Universal Robots URScript: jerry_new_robot_1.script

def Machining2():
  # Default parameters:
  global speed_ms = 0.3
  global speed_rads = 0.75
  global accel_mss = 3
  global accel_radss = 1.2
  global blend_radius_m = 0.001

  # Add subprograms here
  # Start of main program
  # Program generated by RoboDK v5.6.8 for UR10e on 15/12/2023 14:31:05
  # Using nominal kinematics.
  blend_radius_m = 0.001
  speed_ms = 0.01
  # set_reference(p[0.405000, -0.105000, 0.010000, 0.000000, 0.000000, 0.000000])
  set_tcp(p[0.000000, 0.000000, 0.252000, 0.000000, 0.000000, 0.000000])
  # Show Tool
  movej([0.286818, -1.328197, -2.476759, -0.907433, 1.570796, 1.857614],accel_radss,speed_rads,0,blend_radius_m)
  movel([0.286818, -1.380785, -2.509088, -0.822516, 1.570796, 1.857614],accel_mss,speed_ms,0,blend_radius_m)
  speed_ms = 0.01
  movel([0.286818, -1.403946, -2.521184, -0.787258, 1.570796, 1.857614],accel_mss,speed_ms,0,blend_radius_m)
  speed_ms = 0.003
  movel([0.286818, -1.412952, -2.525590, -0.773847, 1.570796, 1.857614],accel_mss,speed_ms,0,blend_radius_m)
  speed_ms = 0.007
  movel([0.278957, -1.415271, -2.523827, -0.773292, 1.570796, 1.849754],accel_mss,speed_ms,0,blend_radius_m)
  movel([0.277121, -1.413155, -2.525436, -0.773798, 1.570796, 1.847918],accel_mss,speed_ms,0,blend_radius_m)
  movel([0.275274, -1.411040, -2.527038, -0.774311, 1.570796, 1.846071],accel_mss,speed_ms,0,blend_radius_m)
  movel([0.275922, -1.409907, -2.527894, -0.774588, 1.570796, 1.846719],accel_mss,speed_ms,0,blend_radius_m)
  movel([0.276572, -1.408773, -2.528749, -0.774868, 1.570796, 1.847368],accel_mss,speed_ms,0,blend_radius_m)
  movel([0.275763, -1.408648, -2.528842, -0.774898, 1.570796, 1.846559],accel_mss,speed_ms,0,blend_radius_m)
  movel([0.268969, -1.407825, -2.529461, -0.775102, 1.570796, 1.839766],accel_mss,speed_ms,0,blend_radius_m)
  movel([0.266583, -1.407546, -2.529671, -0.775172, 1.570796, 1.837380],accel_mss,speed_ms,0,blend_radius_m)
  movel([0.265501, -1.407413, -2.529771, -0.775205, 1.570796, 1.836297],accel_mss,speed_ms,0,blend_radius_m)
  movel([0.264422, -1.407272, -2.529877, -0.775240, 1.570796, 1.835218],accel_mss,speed_ms,0,blend_radius_m)
  movel([0.263348, -1.407121, -2.529990, -0.775278, 1.570796, 1.834144],accel_mss,speed_ms,0,blend_radius_m)
  movel([0.262516, -1.406998, -2.530083, -0.775309, 1.570796, 1.833312],accel_mss,speed_ms,0,blend_radius_m)
  movel([0.261691, -1.406866, -2.530182, -0.775342, 1.570796, 1.832487],accel_mss,speed_ms,0,blend_radius_m)
  movel([0.260873, -1.406721, -2.530290, -0.775378, 1.570796, 1.831670],accel_mss,speed_ms,0,blend_radius_m)
  movel([0.260123, -1.406582, -2.530395, -0.775413, 1.570796, 1.830919],accel_mss,speed_ms,0,blend_radius_m)
  movel([0.259383, -1.406429, -2.530509, -0.775451, 1.570796, 1.830179],accel_mss,speed_ms,0,blend_radius_m)
  movel([0.258650, -1.406263, -2.530633, -0.775493, 1.570796, 1.829447],accel_mss,speed_ms,0,blend_radius_m)
  movel([0.257946, -1.406092, -2.530761, -0.775535, 1.570796, 1.828742],accel_mss,speed_ms,0,blend_radius_m)
  movel([0.257255, -1.405904, -2.530902, -0.775583, 1.570796, 1.828051],accel_mss,speed_ms,0,blend_radius_m)
  movel([0.256572, -1.405700, -2.531055, -0.775634, 1.570796, 1.827368],accel_mss,speed_ms,0,blend_radius_m)
  movel([0.255900, -1.405481, -2.531218, -0.775689, 1.570796, 1.826696],accel_mss,speed_ms,0,blend_radius_m)
  movel([0.255241, -1.405247, -2.531394, -0.775748, 1.570796, 1.826037],accel_mss,speed_ms,0,blend_radius_m)
  movel([0.254785, -1.405071, -2.531525, -0.775793, 1.570796, 1.825581],accel_mss,speed_ms,0,blend_radius_m)
  movel([0.254341, -1.404877, -2.531670, -0.775842, 1.570796, 1.825137],accel_mss,speed_ms,0,blend_radius_m)
  movel([0.253906, -1.404672, -2.531824, -0.775894, 1.570796, 1.824702],accel_mss,speed_ms,0,blend_radius_m)
  movel([0.253487, -1.404450, -2.531989, -0.775950, 1.570796, 1.824283],accel_mss,speed_ms,0,blend_radius_m)
  movel([0.253079, -1.404213, -2.532166, -0.776010, 1.570796, 1.823875],accel_mss,speed_ms,0,blend_radius_m)
  movel([0.252685, -1.403964, -2.532352, -0.776073, 1.570796, 1.823481],accel_mss,speed_ms,0,blend_radius_m)
  movel([0.252356, -1.403735, -2.532523, -0.776131, 1.570796, 1.823152],accel_mss,speed_ms,0,blend_radius_m)
  movel([0.252040, -1.403492, -2.532704, -0.776193, 1.570796, 1.822837],accel_mss,speed_ms,0,blend_radius_m)
  movel([0.251741, -1.403234, -2.532896, -0.776259, 1.570796, 1.822538],accel_mss,speed_ms,0,blend_radius_m)
  movel([0.251455, -1.402963, -2.533098, -0.776328, 1.570796, 1.822252],accel_mss,speed_ms,0,blend_radius_m)
  movel([0.251184, -1.402679, -2.533309, -0.776401, 1.570796, 1.821980],accel_mss,speed_ms,0,blend_radius_m)
  movel([0.250929, -1.402382, -2.533530, -0.776477, 1.570796, 1.821725],accel_mss,speed_ms,0,blend_radius_m)
  movel([0.250744, -1.402139, -2.533711, -0.776540, 1.570796, 1.821540],accel_mss,speed_ms,0,blend_radius_m)
  movel([0.250570, -1.401887, -2.533898, -0.776604, 1.570796, 1.821366],accel_mss,speed_ms,0,blend_radius_m)
  movel([0.250413, -1.401623, -2.534094, -0.776672, 1.570796, 1.821209],accel_mss,speed_ms,0,blend_radius_m)
  movel([0.250269, -1.401348, -2.534298, -0.776743, 1.570796, 1.821066],accel_mss,speed_ms,0,blend_radius_m)
  movel([0.250142, -1.401063, -2.534509, -0.776817, 1.570796, 1.820938],accel_mss,speed_ms,0,blend_radius_m)
  movel([0.250030, -1.400772, -2.534725, -0.776892, 1.570796, 1.820826],accel_mss,speed_ms,0,blend_radius_m)
  movel([0.249933, -1.400468, -2.534950, -0.776970, 1.570796, 1.820729],accel_mss,speed_ms,0,blend_radius_m)
  movel([0.249858, -1.400178, -2.535165, -0.777046, 1.570796, 1.820655],accel_mss,speed_ms,0,blend_radius_m)
  movel([0.249800, -1.399877, -2.535388, -0.777124, 1.570796, 1.820596],accel_mss,speed_ms,0,blend_radius_m)
  movel([0.249762, -1.399567, -2.535617, -0.777205, 1.570796, 1.820559],accel_mss,speed_ms,0,blend_radius_m)
  movel([0.249742, -1.399250, -2.535851, -0.777287, 1.570796, 1.820538],accel_mss,speed_ms,0,blend_radius_m)
  movel([0.249739, -1.398896, -2.536113, -0.777380, 1.570796, 1.820535],accel_mss,speed_ms,0,blend_radius_m)
  movel([0.249750, -1.398537, -2.536378, -0.777474, 1.570796, 1.820546],accel_mss,speed_ms,0,blend_radius_m)
  movel([0.249777, -1.398172, -2.536647, -0.777570, 1.570796, 1.820573],accel_mss,speed_ms,0,blend_radius_m)
  movel([0.249818, -1.397802, -2.536920, -0.777667, 1.570796, 1.820614],accel_mss,speed_ms,0,blend_radius_m)
  movel([0.249880, -1.397415, -2.537205, -0.777769, 1.570796, 1.820676],accel_mss,speed_ms,0,blend_radius_m)
  movel([0.249952, -1.397029, -2.537490, -0.777871, 1.570796, 1.820749],accel_mss,speed_ms,0,blend_radius_m)
  movel([0.250043, -1.396635, -2.537779, -0.777975, 1.570796, 1.820839],accel_mss,speed_ms,0,blend_radius_m)
  movel([0.250147, -1.396242, -2.538068, -0.778079, 1.570796, 1.820943],accel_mss,speed_ms,0,blend_radius_m)
  movel([0.250264, -1.395857, -2.538351, -0.778181, 1.570796, 1.821061],accel_mss,speed_ms,0,blend_radius_m)
  movel([0.250398, -1.395471, -2.538634, -0.778284, 1.570796, 1.821194],accel_mss,speed_ms,0,blend_radius_m)
  movel([0.250547, -1.395084, -2.538918, -0.778387, 1.570796, 1.821344],accel_mss,speed_ms,0,blend_radius_m)
  movel([0.250711, -1.394696, -2.539203, -0.778491, 1.570796, 1.821507],accel_mss,speed_ms,0,blend_radius_m)
  movel([0.250904, -1.394272, -2.539513, -0.778604, 1.570796, 1.821701],accel_mss,speed_ms,0,blend_radius_m)
  movel([0.251110, -1.393847, -2.539824, -0.778719, 1.570796, 1.821906],accel_mss,speed_ms,0,blend_radius_m)
  movel([0.251326, -1.393423, -2.540133, -0.778832, 1.570796, 1.822123],accel_mss,speed_ms,0,blend_radius_m)
  movel([0.251379, -1.393339, -2.540195, -0.778855, 1.570796, 1.822175],accel_mss,speed_ms,0,blend_radius_m)
  movel([0.251441, -1.393255, -2.540256, -0.778878, 1.570796, 1.822237],accel_mss,speed_ms,0,blend_radius_m)
  movel([0.251514, -1.393178, -2.540313, -0.778899, 1.570796, 1.822310],accel_mss,speed_ms,0,blend_radius_m)
  movel([0.251592, -1.393106, -2.540365, -0.778918, 1.570796, 1.822389],accel_mss,speed_ms,0,blend_radius_m)
  movel([0.251680, -1.393042, -2.540412, -0.778935, 1.570796, 1.822476],accel_mss,speed_ms,0,blend_radius_m)
  movel([0.251772, -1.392987, -2.540452, -0.778950, 1.570796, 1.822568],accel_mss,speed_ms,0,blend_radius_m)
  movel([0.251894, -1.392931, -2.540493, -0.778965, 1.570796, 1.822690],accel_mss,speed_ms,0,blend_radius_m)
  movel([0.252016, -1.392887, -2.540525, -0.778977, 1.570796, 1.822813],accel_mss,speed_ms,0,blend_radius_m)
  movel([0.252140, -1.392857, -2.540547, -0.778985, 1.570796, 1.822936],accel_mss,speed_ms,0,blend_radius_m)
  movel([0.252259, -1.392843, -2.540557, -0.778989, 1.570796, 1.823055],accel_mss,speed_ms,0,blend_radius_m)
  movel([0.252371, -1.392844, -2.540556, -0.778989, 1.570796, 1.823167],accel_mss,speed_ms,0,blend_radius_m)
  movel([0.252874, -1.392895, -2.540519, -0.778975, 1.570796, 1.823670],accel_mss,speed_ms,0,blend_radius_m)
  movel([0.253372, -1.392952, -2.540477, -0.778959, 1.570796, 1.824168],accel_mss,speed_ms,0,blend_radius_m)
  movel([0.253866, -1.393017, -2.540430, -0.778942, 1.570796, 1.824662],accel_mss,speed_ms,0,blend_radius_m)
  movel([0.254596, -1.393123, -2.540352, -0.778913, 1.570796, 1.825392],accel_mss,speed_ms,0,blend_radius_m)
  movel([0.254793, -1.392422, -2.540864, -0.779103, 1.570796, 1.825589],accel_mss,speed_ms,0,blend_radius_m)
  movel([0.254989, -1.391722, -2.541374, -0.779293, 1.570796, 1.825785],accel_mss,speed_ms,0,blend_radius_m)
  movel([0.238692, -1.394040, -2.539683, -0.778667, 1.570796, 1.809488],accel_mss,speed_ms,0,blend_radius_m)
  movel([0.229160, -1.395492, -2.538618, -0.778278, 1.570796, 1.799956],accel_mss,speed_ms,0,blend_radius_m)
  movel([0.227094, -1.395812, -2.538384, -0.778193, 1.570796, 1.797890],accel_mss,speed_ms,0,blend_radius_m)
  movel([0.225031, -1.396124, -2.538155, -0.778110, 1.570796, 1.795827],accel_mss,speed_ms,0,blend_radius_m)
  movel([0.222484, -1.396503, -2.537876, -0.778010, 1.570796, 1.793281],accel_mss,speed_ms,0,blend_radius_m)
  movel([0.222392, -1.396509, -2.537872, -0.778008, 1.570796, 1.793189],accel_mss,speed_ms,0,blend_radius_m)
  movel([0.222306, -1.396503, -2.537876, -0.778010, 1.570796, 1.793102],accel_mss,speed_ms,0,blend_radius_m)
  movel([0.222225, -1.396485, -2.537890, -0.778014, 1.570796, 1.793021],accel_mss,speed_ms,0,blend_radius_m)
  movel([0.222156, -1.396453, -2.537913, -0.778023, 1.570796, 1.792952],accel_mss,speed_ms,0,blend_radius_m)
  movel([0.222108, -1.396419, -2.537938, -0.778032, 1.570796, 1.792904],accel_mss,speed_ms,0,blend_radius_m)
  movel([0.222070, -1.396378, -2.537968, -0.778043, 1.570796, 1.792867],accel_mss,speed_ms,0,blend_radius_m)
  movel([0.222044, -1.396328, -2.538005, -0.778056, 1.570796, 1.792841],accel_mss,speed_ms,0,blend_radius_m)
  movel([0.222025, -1.396269, -2.538048, -0.778072, 1.570796, 1.792821],accel_mss,speed_ms,0,blend_radius_m)
  movel([0.222016, -1.396204, -2.538096, -0.778089, 1.570796, 1.792812],accel_mss,speed_ms,0,blend_radius_m)
  movel([0.222016, -1.396138, -2.538144, -0.778106, 1.570796, 1.792813],accel_mss,speed_ms,0,blend_radius_m)
  movel([0.222040, -1.395960, -2.538275, -0.778154, 1.570796, 1.792836],accel_mss,speed_ms,0,blend_radius_m)
  movel([0.222075, -1.395781, -2.538407, -0.778201, 1.570796, 1.792872],accel_mss,speed_ms,0,blend_radius_m)
  movel([0.222291, -1.394877, -2.539069, -0.778442, 1.570796, 1.793087],accel_mss,speed_ms,0,blend_radius_m)
  movel([0.222650, -1.393424, -2.540133, -0.778832, 1.570796, 1.793446],accel_mss,speed_ms,0,blend_radius_m)
  movel([0.212968, -1.395043, -2.538948, -0.778398, 1.570796, 1.783765],accel_mss,speed_ms,0,blend_radius_m)
  movel([0.203286, -1.396738, -2.537704, -0.777948, 1.570796, 1.774082],accel_mss,speed_ms,0,blend_radius_m)
  movel([0.203152, -1.397328, -2.537269, -0.777792, 1.570796, 1.773949],accel_mss,speed_ms,0,blend_radius_m)
  movel([0.203019, -1.397918, -2.536835, -0.777636, 1.570796, 1.773815],accel_mss,speed_ms,0,blend_radius_m)
  movel([0.186235, -1.401026, -2.534537, -0.776826, 1.570796, 1.757031],accel_mss,speed_ms,0,blend_radius_m)
  movel([0.169460, -1.404353, -2.532062, -0.775974, 1.570796, 1.740256],accel_mss,speed_ms,0,blend_radius_m)
  movel([0.168502, -1.404999, -2.531579, -0.775811, 1.570796, 1.739298],accel_mss,speed_ms,0,blend_radius_m)
  movel([0.168210, -1.405190, -2.531436, -0.775763, 1.570796, 1.739006],accel_mss,speed_ms,0,blend_radius_m)
  movel([0.167917, -1.405378, -2.531296, -0.775715, 1.570796, 1.738713],accel_mss,speed_ms,0,blend_radius_m)
  movel([0.167618, -1.405559, -2.531161, -0.775670, 1.570796, 1.738414],accel_mss,speed_ms,0,blend_radius_m)
  movel([0.167135, -1.405842, -2.530948, -0.775598, 1.570796, 1.737931],accel_mss,speed_ms,0,blend_radius_m)
  movel([0.166648, -1.406110, -2.530748, -0.775531, 1.570796, 1.737444],accel_mss,speed_ms,0,blend_radius_m)
  movel([0.166146, -1.406376, -2.530549, -0.775464, 1.570796, 1.736942],accel_mss,speed_ms,0,blend_radius_m)
  movel([0.165641, -1.406626, -2.530362, -0.775402, 1.570796, 1.736437],accel_mss,speed_ms,0,blend_radius_m)
  movel([0.165143, -1.406860, -2.530186, -0.775343, 1.570796, 1.735939],accel_mss,speed_ms,0,blend_radius_m)
  movel([0.164644, -1.407079, -2.530022, -0.775288, 1.570796, 1.735440],accel_mss,speed_ms,0,blend_radius_m)
  movel([0.164316, -1.407211, -2.529922, -0.775255, 1.570796, 1.735113],accel_mss,speed_ms,0,blend_radius_m)
  movel([0.163987, -1.407330, -2.529833, -0.775226, 1.570796, 1.734783],accel_mss,speed_ms,0,blend_radius_m)
  movel([0.163661, -1.407432, -2.529756, -0.775200, 1.570796, 1.734457],accel_mss,speed_ms,0,blend_radius_m)
  movel([0.162882, -1.407653, -2.529590, -0.775145, 1.570796, 1.733678],accel_mss,speed_ms,0,blend_radius_m)
  movel([0.162106, -1.407860, -2.529435, -0.775094, 1.570796, 1.732902],accel_mss,speed_ms,0,blend_radius_m)
  movel([0.161310, -1.408059, -2.529285, -0.775044, 1.570796, 1.732107],accel_mss,speed_ms,0,blend_radius_m)
  movel([0.160517, -1.408252, -2.529140, -0.774996, 1.570796, 1.731313],accel_mss,speed_ms,0,blend_radius_m)
  movel([0.160414, -1.408270, -2.529127, -0.774992, 1.570796, 1.731210],accel_mss,speed_ms,0,blend_radius_m)
  movel([0.160319, -1.408272, -2.529125, -0.774992, 1.570796, 1.731115],accel_mss,speed_ms,0,blend_radius_m)
  movel([0.160228, -1.408261, -2.529134, -0.774994, 1.570796, 1.731025],accel_mss,speed_ms,0,blend_radius_m)
  movel([0.160150, -1.408233, -2.529155, -0.775001, 1.570796, 1.730946],accel_mss,speed_ms,0,blend_radius_m)
  movel([0.160120, -1.408213, -2.529170, -0.775006, 1.570796, 1.730916],accel_mss,speed_ms,0,blend_radius_m)
  movel([0.160100, -1.408185, -2.529191, -0.775013, 1.570796, 1.730896],accel_mss,speed_ms,0,blend_radius_m)
  movel([0.160090, -1.408151, -2.529216, -0.775021, 1.570796, 1.730887],accel_mss,speed_ms,0,blend_radius_m)
  movel([0.160090, -1.408113, -2.529245, -0.775031, 1.570796, 1.730887],accel_mss,speed_ms,0,blend_radius_m)
  movel([0.160497, -1.405621, -2.531114, -0.775654, 1.570796, 1.731293],accel_mss,speed_ms,0,blend_radius_m)
  movel([0.160790, -1.403859, -2.532430, -0.776100, 1.570796, 1.731586],accel_mss,speed_ms,0,blend_radius_m)
  movel([0.161094, -1.402089, -2.533748, -0.776552, 1.570796, 1.731890],accel_mss,speed_ms,0,blend_radius_m)
  movel([0.162202, -1.395764, -2.538419, -0.778206, 1.570796, 1.732999],accel_mss,speed_ms,0,blend_radius_m)
  movel([0.164448, -1.383126, -2.547582, -0.781681, 1.570796, 1.735244],accel_mss,speed_ms,0,blend_radius_m)
  movel([0.164830, -1.383043, -2.547641, -0.781705, 1.570796, 1.735626],accel_mss,speed_ms,0,blend_radius_m)
  movel([0.165050, -1.382984, -2.547683, -0.781721, 1.570796, 1.735846],accel_mss,speed_ms,0,blend_radius_m)
  movel([0.165159, -1.382921, -2.547729, -0.781739, 1.570796, 1.735955],accel_mss,speed_ms,0,blend_radius_m)
  movel([0.165225, -1.382825, -2.547797, -0.781767, 1.570796, 1.736022],accel_mss,speed_ms,0,blend_radius_m)
  movel([0.165270, -1.382649, -2.547923, -0.781817, 1.570796, 1.736066],accel_mss,speed_ms,0,blend_radius_m)
  movel([0.165294, -1.382556, -2.547990, -0.781843, 1.570796, 1.736090],accel_mss,speed_ms,0,blend_radius_m)
  movel([0.165328, -1.382461, -2.548058, -0.781870, 1.570796, 1.736124],accel_mss,speed_ms,0,blend_radius_m)
  movel([0.165349, -1.382421, -2.548086, -0.781882, 1.570796, 1.736145],accel_mss,speed_ms,0,blend_radius_m)
  movel([0.165379, -1.382383, -2.548113, -0.781893, 1.570796, 1.736176],accel_mss,speed_ms,0,blend_radius_m)
  movel([0.165418, -1.382352, -2.548136, -0.781902, 1.570796, 1.736214],accel_mss,speed_ms,0,blend_radius_m)
  movel([0.165499, -1.382303, -2.548171, -0.781915, 1.570796, 1.736295],accel_mss,speed_ms,0,blend_radius_m)
  movel([0.165585, -1.382265, -2.548198, -0.781926, 1.570796, 1.736381],accel_mss,speed_ms,0,blend_radius_m)
  movel([0.166012, -1.382128, -2.548296, -0.781965, 1.570796, 1.736808],accel_mss,speed_ms,0,blend_radius_m)
  movel([0.166274, -1.382054, -2.548348, -0.781986, 1.570796, 1.737070],accel_mss,speed_ms,0,blend_radius_m)
  movel([0.166534, -1.381992, -2.548393, -0.782004, 1.570796, 1.737330],accel_mss,speed_ms,0,blend_radius_m)
  movel([0.166792, -1.381940, -2.548430, -0.782019, 1.570796, 1.737589],accel_mss,speed_ms,0,blend_radius_m)
  movel([0.167305, -1.381853, -2.548492, -0.782044, 1.570796, 1.738102],accel_mss,speed_ms,0,blend_radius_m)
  movel([0.167813, -1.381783, -2.548542, -0.782064, 1.570796, 1.738609],accel_mss,speed_ms,0,blend_radius_m)
  movel([0.168346, -1.381724, -2.548584, -0.782081, 1.570796, 1.739143],accel_mss,speed_ms,0,blend_radius_m)
  movel([0.168877, -1.381683, -2.548614, -0.782092, 1.570796, 1.739673],accel_mss,speed_ms,0,blend_radius_m)
  movel([0.169191, -1.381665, -2.548626, -0.782098, 1.570796, 1.739987],accel_mss,speed_ms,0,blend_radius_m)
  movel([0.169501, -1.381659, -2.548631, -0.782099, 1.570796, 1.740297],accel_mss,speed_ms,0,blend_radius_m)
  movel([0.169807, -1.381660, -2.548630, -0.782099, 1.570796, 1.740603],accel_mss,speed_ms,0,blend_radius_m)
  movel([0.170079, -1.381669, -2.548624, -0.782097, 1.570796, 1.740875],accel_mss,speed_ms,0,blend_radius_m)
  movel([0.170344, -1.381689, -2.548609, -0.782091, 1.570796, 1.741141],accel_mss,speed_ms,0,blend_radius_m)
  movel([0.170606, -1.381717, -2.548590, -0.782083, 1.570796, 1.741402],accel_mss,speed_ms,0,blend_radius_m)
  movel([0.171068, -1.381785, -2.548541, -0.782063, 1.570796, 1.741865],accel_mss,speed_ms,0,blend_radius_m)
  movel([0.171524, -1.381865, -2.548483, -0.782040, 1.570796, 1.742320],accel_mss,speed_ms,0,blend_radius_m)
  movel([0.171974, -1.381962, -2.548415, -0.782013, 1.570796, 1.742770],accel_mss,speed_ms,0,blend_radius_m)
  movel([0.172412, -1.382071, -2.548336, -0.781982, 1.570796, 1.743208],accel_mss,speed_ms,0,blend_radius_m)
  movel([0.172651, -1.382141, -2.548286, -0.781961, 1.570796, 1.743447],accel_mss,speed_ms,0,blend_radius_m)
  movel([0.172886, -1.382221, -2.548229, -0.781939, 1.570796, 1.743682],accel_mss,speed_ms,0,blend_radius_m)
  movel([0.173112, -1.382309, -2.548166, -0.781914, 1.570796, 1.743908],accel_mss,speed_ms,0,blend_radius_m)
  movel([0.173605, -1.382514, -2.548020, -0.781855, 1.570796, 1.744401],accel_mss,speed_ms,0,blend_radius_m)
  movel([0.190906, -1.378978, -2.550540, -0.782871, 1.570796, 1.761702],accel_mss,speed_ms,0,blend_radius_m)
  movel([0.208219, -1.375672, -2.552880, -0.783837, 1.570796, 1.779015],accel_mss,speed_ms,0,blend_radius_m)
  movel([0.208066, -1.376337, -2.552411, -0.783642, 1.570796, 1.778862],accel_mss,speed_ms,0,blend_radius_m)
  movel([0.207913, -1.377000, -2.551942, -0.783447, 1.570796, 1.778709],accel_mss,speed_ms,0,blend_radius_m)
  movel([0.212684, -1.376133, -2.552555, -0.783702, 1.570796, 1.783480],accel_mss,speed_ms,0,blend_radius_m)
  movel([0.217469, -1.375223, -2.553196, -0.783969, 1.570796, 1.788265],accel_mss,speed_ms,0,blend_radius_m)
  movel([0.217297, -1.374328, -2.553827, -0.784234, 1.570796, 1.788093],accel_mss,speed_ms,0,blend_radius_m)
  movel([0.217253, -1.374069, -2.554009, -0.784311, 1.570796, 1.788049],accel_mss,speed_ms,0,blend_radius_m)
  movel([0.217221, -1.373807, -2.554194, -0.784389, 1.570796, 1.788017],accel_mss,speed_ms,0,blend_radius_m)
  movel([0.217200, -1.373555, -2.554371, -0.784464, 1.570796, 1.787996],accel_mss,speed_ms,0,blend_radius_m)
  movel([0.217190, -1.373298, -2.554551, -0.784540, 1.570796, 1.787986],accel_mss,speed_ms,0,blend_radius_m)
  movel([0.217192, -1.373038, -2.554734, -0.784618, 1.570796, 1.787988],accel_mss,speed_ms,0,blend_radius_m)
  movel([0.217206, -1.372767, -2.554924, -0.784699, 1.570796, 1.788002],accel_mss,speed_ms,0,blend_radius_m)
  movel([0.217230, -1.372493, -2.555115, -0.784780, 1.570796, 1.788026],accel_mss,speed_ms,0,blend_radius_m)
  movel([0.217264, -1.372216, -2.555310, -0.784863, 1.570796, 1.788060],accel_mss,speed_ms,0,blend_radius_m)
  movel([0.217314, -1.371908, -2.555526, -0.784955, 1.570796, 1.788111],accel_mss,speed_ms,0,blend_radius_m)
  movel([0.217375, -1.371598, -2.555742, -0.785048, 1.570796, 1.788171],accel_mss,speed_ms,0,blend_radius_m)
  movel([0.217443, -1.371287, -2.555960, -0.785142, 1.570796, 1.788239],accel_mss,speed_ms,0,blend_radius_m)
  movel([0.217532, -1.370935, -2.556206, -0.785248, 1.570796, 1.788328],accel_mss,speed_ms,0,blend_radius_m)
  movel([0.217633, -1.370581, -2.556453, -0.785354, 1.570796, 1.788429],accel_mss,speed_ms,0,blend_radius_m)
  movel([0.217749, -1.370225, -2.556702, -0.785462, 1.570796, 1.788545],accel_mss,speed_ms,0,blend_radius_m)
  movel([0.217869, -1.369901, -2.556928, -0.785560, 1.570796, 1.788665],accel_mss,speed_ms,0,blend_radius_m)
  movel([0.218003, -1.369575, -2.557155, -0.785658, 1.570796, 1.788799],accel_mss,speed_ms,0,blend_radius_m)
  movel([0.218156, -1.369250, -2.557382, -0.785757, 1.570796, 1.788952],accel_mss,speed_ms,0,blend_radius_m)
  movel([0.218328, -1.368913, -2.557617, -0.785859, 1.570796, 1.789124],accel_mss,speed_ms,0,blend_radius_m)
  movel([0.218513, -1.368579, -2.557849, -0.785961, 1.570796, 1.789309],accel_mss,speed_ms,0,blend_radius_m)
  movel([0.218715, -1.368245, -2.558082, -0.786063, 1.570796, 1.789511],accel_mss,speed_ms,0,blend_radius_m)
  movel([0.218964, -1.367856, -2.558351, -0.786181, 1.570796, 1.789761],accel_mss,speed_ms,0,blend_radius_m)
  movel([0.219223, -1.367471, -2.558619, -0.786299, 1.570796, 1.790019],accel_mss,speed_ms,0,blend_radius_m)
  movel([0.219493, -1.367087, -2.558885, -0.786417, 1.570796, 1.790290],accel_mss,speed_ms,0,blend_radius_m)
  movel([0.220268, -1.366008, -2.559633, -0.786748, 1.570796, 1.791064],accel_mss,speed_ms,0,blend_radius_m)
  movel([0.218931, -1.366247, -2.559468, -0.786674, 1.570796, 1.789727],accel_mss,speed_ms,0,blend_radius_m)
  movel([0.217591, -1.366488, -2.559301, -0.786601, 1.570796, 1.788387],accel_mss,speed_ms,0,blend_radius_m)
  movel([0.217739, -1.365869, -2.559729, -0.786791, 1.570796, 1.788535],accel_mss,speed_ms,0,blend_radius_m)
  movel([0.217888, -1.365249, -2.560158, -0.786982, 1.570796, 1.788684],accel_mss,speed_ms,0,blend_radius_m)
  movel([0.213855, -1.365983, -2.559650, -0.786756, 1.570796, 1.784651],accel_mss,speed_ms,0,blend_radius_m)
  movel([0.209822, -1.366730, -2.559133, -0.786526, 1.570796, 1.780618],accel_mss,speed_ms,0,blend_radius_m)
  movel([0.209666, -1.367404, -2.558666, -0.786320, 1.570796, 1.780462],accel_mss,speed_ms,0,blend_radius_m)
  movel([0.209510, -1.368076, -2.558199, -0.786114, 1.570796, 1.780306],accel_mss,speed_ms,0,blend_radius_m)
  movel([0.191959, -1.371470, -2.555832, -0.785087, 1.570796, 1.762755],accel_mss,speed_ms,0,blend_radius_m)
  movel([0.174421, -1.375101, -2.553282, -0.784005, 1.570796, 1.745218],accel_mss,speed_ms,0,blend_radius_m)
  movel([0.173235, -1.375825, -2.552772, -0.783792, 1.570796, 1.744031],accel_mss,speed_ms,0,blend_radius_m)
  movel([0.172826, -1.376067, -2.552601, -0.783721, 1.570796, 1.743622],accel_mss,speed_ms,0,blend_radius_m)
  movel([0.172415, -1.376300, -2.552436, -0.783652, 1.570796, 1.743211],accel_mss,speed_ms,0,blend_radius_m)
  movel([0.172001, -1.376524, -2.552278, -0.783587, 1.570796, 1.742797],accel_mss,speed_ms,0,blend_radius_m)
  movel([0.171584, -1.376736, -2.552129, -0.783525, 1.570796, 1.742381],accel_mss,speed_ms,0,blend_radius_m)
  movel([0.171160, -1.376943, -2.551982, -0.783464, 1.570796, 1.741956],accel_mss,speed_ms,0,blend_radius_m)
  movel([0.170730, -1.377139, -2.551844, -0.783407, 1.570796, 1.741527],accel_mss,speed_ms,0,blend_radius_m)
  movel([0.170303, -1.377326, -2.551711, -0.783352, 1.570796, 1.741099],accel_mss,speed_ms,0,blend_radius_m)
  movel([0.169873, -1.377501, -2.551587, -0.783301, 1.570796, 1.740670],accel_mss,speed_ms,0,blend_radius_m)
  movel([0.169451, -1.377661, -2.551474, -0.783254, 1.570796, 1.740247],accel_mss,speed_ms,0,blend_radius_m)
  movel([0.169028, -1.377814, -2.551365, -0.783210, 1.570796, 1.739824],accel_mss,speed_ms,0,blend_radius_m)
  movel([0.168605, -1.377954, -2.551266, -0.783169, 1.570796, 1.739402],accel_mss,speed_ms,0,blend_radius_m)
  movel([0.168183, -1.378082, -2.551176, -0.783131, 1.570796, 1.738979],accel_mss,speed_ms,0,blend_radius_m)
  movel([0.167784, -1.378194, -2.551096, -0.783099, 1.570796, 1.738580],accel_mss,speed_ms,0,blend_radius_m)
  movel([0.167388, -1.378291, -2.551027, -0.783071, 1.570796, 1.738184],accel_mss,speed_ms,0,blend_radius_m)
  movel([0.166994, -1.378377, -2.550966, -0.783046, 1.570796, 1.737791],accel_mss,speed_ms,0,blend_radius_m)
  movel([0.166604, -1.378448, -2.550916, -0.783025, 1.570796, 1.737400],accel_mss,speed_ms,0,blend_radius_m)
  movel([0.166192, -1.378515, -2.550869, -0.783006, 1.570796, 1.736989],accel_mss,speed_ms,0,blend_radius_m)
  movel([0.165843, -1.378566, -2.550832, -0.782991, 1.570796, 1.736639],accel_mss,speed_ms,0,blend_radius_m)
  movel([0.165544, -1.378607, -2.550803, -0.782979, 1.570796, 1.736340],accel_mss,speed_ms,0,blend_radius_m)
  movel([0.165523, -1.378605, -2.550804, -0.782979, 1.570796, 1.736319],accel_mss,speed_ms,0,blend_radius_m)
  movel([0.165508, -1.378598, -2.550809, -0.782981, 1.570796, 1.736304],accel_mss,speed_ms,0,blend_radius_m)
  movel([0.165499, -1.378581, -2.550822, -0.782986, 1.570796, 1.736296],accel_mss,speed_ms,0,blend_radius_m)
  movel([0.165498, -1.378562, -2.550835, -0.782992, 1.570796, 1.736295],accel_mss,speed_ms,0,blend_radius_m)
  movel([0.166175, -1.374788, -2.553503, -0.784098, 1.570796, 1.736971],accel_mss,speed_ms,0,blend_radius_m)
  movel([0.166934, -1.370595, -2.556444, -0.785350, 1.570796, 1.737730],accel_mss,speed_ms,0,blend_radius_m)
  movel([0.167851, -1.365586, -2.559925, -0.786878, 1.570796, 1.738647],accel_mss,speed_ms,0,blend_radius_m)
  movel([0.170300, -1.352354, -2.568954, -0.791082, 1.570796, 1.741096],accel_mss,speed_ms,0,blend_radius_m)
  movel([0.170708, -1.352260, -2.569016, -0.791112, 1.570796, 1.741504],accel_mss,speed_ms,0,blend_radius_m)
  movel([0.171055, -1.352136, -2.569100, -0.791153, 1.570796, 1.741852],accel_mss,speed_ms,0,blend_radius_m)
  movel([0.171088, -1.352091, -2.569130, -0.791167, 1.570796, 1.741884],accel_mss,speed_ms,0,blend_radius_m)
  movel([0.171101, -1.352045, -2.569162, -0.791183, 1.570796, 1.741898],accel_mss,speed_ms,0,blend_radius_m)
  movel([0.171107, -1.351852, -2.569291, -0.791246, 1.570796, 1.741903],accel_mss,speed_ms,0,blend_radius_m)
  movel([0.171108, -1.351756, -2.569356, -0.791277, 1.570796, 1.741905],accel_mss,speed_ms,0,blend_radius_m)
  movel([0.171118, -1.351656, -2.569423, -0.791310, 1.570796, 1.741914],accel_mss,speed_ms,0,blend_radius_m)
  movel([0.171127, -1.351619, -2.569448, -0.791322, 1.570796, 1.741924],accel_mss,speed_ms,0,blend_radius_m)
  movel([0.171151, -1.351583, -2.569472, -0.791334, 1.570796, 1.741947],accel_mss,speed_ms,0,blend_radius_m)
  movel([0.171181, -1.351550, -2.569494, -0.791345, 1.570796, 1.741977],accel_mss,speed_ms,0,blend_radius_m)
  movel([0.171246, -1.351501, -2.569528, -0.791361, 1.570796, 1.742042],accel_mss,speed_ms,0,blend_radius_m)
  movel([0.171317, -1.351465, -2.569552, -0.791373, 1.570796, 1.742114],accel_mss,speed_ms,0,blend_radius_m)
  movel([0.171697, -1.351324, -2.569646, -0.791419, 1.570796, 1.742493],accel_mss,speed_ms,0,blend_radius_m)
  movel([0.171915, -1.351250, -2.569696, -0.791443, 1.570796, 1.742711],accel_mss,speed_ms,0,blend_radius_m)
  movel([0.172130, -1.351190, -2.569736, -0.791463, 1.570796, 1.742926],accel_mss,speed_ms,0,blend_radius_m)
  movel([0.172344, -1.351140, -2.569770, -0.791479, 1.570796, 1.743140],accel_mss,speed_ms,0,blend_radius_m)
  movel([0.172800, -1.351049, -2.569831, -0.791509, 1.570796, 1.743596],accel_mss,speed_ms,0,blend_radius_m)
  movel([0.173254, -1.350971, -2.569884, -0.791535, 1.570796, 1.744051],accel_mss,speed_ms,0,blend_radius_m)
  movel([0.173743, -1.350899, -2.569931, -0.791558, 1.570796, 1.744539],accel_mss,speed_ms,0,blend_radius_m)
  movel([0.174229, -1.350840, -2.569971, -0.791578, 1.570796, 1.745026],accel_mss,speed_ms,0,blend_radius_m)
  movel([0.174671, -1.350801, -2.569997, -0.791591, 1.570796, 1.745467],accel_mss,speed_ms,0,blend_radius_m)
  movel([0.175104, -1.350780, -2.570011, -0.791598, 1.570796, 1.745901],accel_mss,speed_ms,0,blend_radius_m)
  movel([0.175523, -1.350771, -2.570018, -0.791601, 1.570796, 1.746320],accel_mss,speed_ms,0,blend_radius_m)
  movel([0.175932, -1.350777, -2.570013, -0.791598, 1.570796, 1.746729],accel_mss,speed_ms,0,blend_radius_m)
  movel([0.176336, -1.350796, -2.570001, -0.791592, 1.570796, 1.747133],accel_mss,speed_ms,0,blend_radius_m)
  movel([0.176721, -1.350828, -2.569979, -0.791582, 1.570796, 1.747517],accel_mss,speed_ms,0,blend_radius_m)
  movel([0.177098, -1.350872, -2.569950, -0.791567, 1.570796, 1.747894],accel_mss,speed_ms,0,blend_radius_m)
  movel([0.177467, -1.350932, -2.569910, -0.791548, 1.570796, 1.748264],accel_mss,speed_ms,0,blend_radius_m)
  movel([0.177834, -1.351005, -2.569860, -0.791524, 1.570796, 1.748630],accel_mss,speed_ms,0,blend_radius_m)
  movel([0.178187, -1.351094, -2.569800, -0.791494, 1.570796, 1.748984],accel_mss,speed_ms,0,blend_radius_m)
  movel([0.178536, -1.351196, -2.569732, -0.791461, 1.570796, 1.749333],accel_mss,speed_ms,0,blend_radius_m)
  movel([0.178893, -1.351315, -2.569652, -0.791422, 1.570796, 1.749690],accel_mss,speed_ms,0,blend_radius_m)
  movel([0.179243, -1.351447, -2.569563, -0.791378, 1.570796, 1.750039],accel_mss,speed_ms,0,blend_radius_m)
  movel([0.179583, -1.351592, -2.569466, -0.791331, 1.570796, 1.750379],accel_mss,speed_ms,0,blend_radius_m)
  movel([0.180373, -1.351948, -2.569227, -0.791214, 1.570796, 1.751169],accel_mss,speed_ms,0,blend_radius_m)
  movel([0.197715, -1.348255, -2.571701, -0.792432, 1.570796, 1.768511],accel_mss,speed_ms,0,blend_radius_m)
  movel([0.215070, -1.344794, -2.574004, -0.793591, 1.570796, 1.785866],accel_mss,speed_ms,0,blend_radius_m)
  movel([0.214837, -1.345782, -2.573348, -0.793258, 1.570796, 1.785633],accel_mss,speed_ms,0,blend_radius_m)
  movel([0.214678, -1.346640, -2.572778, -0.792971, 1.570796, 1.785474],accel_mss,speed_ms,0,blend_radius_m)
  movel([0.214695, -1.346707, -2.572733, -0.792948, 1.570796, 1.785492],accel_mss,speed_ms,0,blend_radius_m)
  movel([0.214739, -1.346756, -2.572701, -0.792932, 1.570796, 1.785535],accel_mss,speed_ms,0,blend_radius_m)
  movel([0.214900, -1.346820, -2.572658, -0.792911, 1.570796, 1.785697],accel_mss,speed_ms,0,blend_radius_m)
  movel([0.215034, -1.346830, -2.572652, -0.792907, 1.570796, 1.785830],accel_mss,speed_ms,0,blend_radius_m)
  movel([0.215178, -1.346816, -2.572661, -0.792912, 1.570796, 1.785975],accel_mss,speed_ms,0,blend_radius_m)
  movel([0.221027, -1.345762, -2.573362, -0.793265, 1.570796, 1.791823],accel_mss,speed_ms,0,blend_radius_m)
  movel([0.235297, -1.343183, -2.575070, -0.794135, 1.570796, 1.806093],accel_mss,speed_ms,0,blend_radius_m)
  movel([0.235768, -1.341349, -2.576280, -0.794760, 1.570796, 1.806564],accel_mss,speed_ms,0,blend_radius_m)
  movel([0.236034, -1.340342, -2.576942, -0.795104, 1.570796, 1.806830],accel_mss,speed_ms,0,blend_radius_m)
  movel([0.236112, -1.340075, -2.577117, -0.795196, 1.570796, 1.806908],accel_mss,speed_ms,0,blend_radius_m)
  movel([0.236203, -1.339806, -2.577294, -0.795289, 1.570796, 1.806999],accel_mss,speed_ms,0,blend_radius_m)
  movel([0.236268, -1.339638, -2.577405, -0.795347, 1.570796, 1.807064],accel_mss,speed_ms,0,blend_radius_m)
  movel([0.236346, -1.339471, -2.577514, -0.795404, 1.570796, 1.807143],accel_mss,speed_ms,0,blend_radius_m)
  movel([0.236389, -1.339399, -2.577561, -0.795429, 1.570796, 1.807185],accel_mss,speed_ms,0,blend_radius_m)
  movel([0.236441, -1.339327, -2.577609, -0.795454, 1.570796, 1.807237],accel_mss,speed_ms,0,blend_radius_m)
  movel([0.236504, -1.339260, -2.577653, -0.795477, 1.570796, 1.807300],accel_mss,speed_ms,0,blend_radius_m)
  movel([0.236589, -1.339189, -2.577699, -0.795501, 1.570796, 1.807386],accel_mss,speed_ms,0,blend_radius_m)
  movel([0.236684, -1.339129, -2.577738, -0.795522, 1.570796, 1.807480],accel_mss,speed_ms,0,blend_radius_m)
  movel([0.236781, -1.339085, -2.577767, -0.795537, 1.570796, 1.807577],accel_mss,speed_ms,0,blend_radius_m)
  movel([0.236877, -1.339057, -2.577785, -0.795547, 1.570796, 1.807673],accel_mss,speed_ms,0,blend_radius_m)
  movel([0.238008, -1.338836, -2.577930, -0.795623, 1.570796, 1.808804],accel_mss,speed_ms,0,blend_radius_m)
  movel([0.239139, -1.338623, -2.578070, -0.795696, 1.570796, 1.809935],accel_mss,speed_ms,0,blend_radius_m)
  movel([0.241092, -1.338266, -2.578303, -0.795820, 1.570796, 1.811888],accel_mss,speed_ms,0,blend_radius_m)
  movel([0.243044, -1.337924, -2.578527, -0.795938, 1.570796, 1.813840],accel_mss,speed_ms,0,blend_radius_m)
  movel([0.253938, -1.336105, -2.579714, -0.796570, 1.570796, 1.824734],accel_mss,speed_ms,0,blend_radius_m)
  movel([0.271089, -1.333447, -2.581440, -0.797502, 1.570796, 1.841885],accel_mss,speed_ms,0,blend_radius_m)
  movel([0.271605, -1.331677, -2.582584, -0.798127, 1.570796, 1.842402],accel_mss,speed_ms,0,blend_radius_m)
  movel([0.272125, -1.329900, -2.583729, -0.798760, 1.570796, 1.842921],accel_mss,speed_ms,0,blend_radius_m)
  movel([0.261552, -1.328518, -2.584616, -0.799255, 1.570796, 1.832348],accel_mss,speed_ms,0,blend_radius_m)
  movel([0.250887, -1.327288, -2.585404, -0.799697, 1.570796, 1.821683],accel_mss,speed_ms,0,blend_radius_m)
  movel([0.250851, -1.327305, -2.585393, -0.799691, 1.570796, 1.821647],accel_mss,speed_ms,0,blend_radius_m)
  movel([0.249681, -1.329503, -2.583984, -0.798902, 1.570796, 1.820477],accel_mss,speed_ms,0,blend_radius_m)
  movel([0.245732, -1.330878, -2.583100, -0.798411, 1.570796, 1.816528],accel_mss,speed_ms,0,blend_radius_m)
  movel([0.244205, -1.331410, -2.582757, -0.798222, 1.570796, 1.815002],accel_mss,speed_ms,0,blend_radius_m)
  movel([0.242889, -1.331865, -2.582463, -0.798061, 1.570796, 1.813685],accel_mss,speed_ms,0,blend_radius_m)
  movel([0.241743, -1.332258, -2.582209, -0.797922, 1.570796, 1.812540],accel_mss,speed_ms,0,blend_radius_m)
  movel([0.241668, -1.332280, -2.582195, -0.797914, 1.570796, 1.812464],accel_mss,speed_ms,0,blend_radius_m)
  movel([0.241591, -1.332296, -2.582185, -0.797908, 1.570796, 1.812388],accel_mss,speed_ms,0,blend_radius_m)
  movel([0.241512, -1.332305, -2.582179, -0.797905, 1.570796, 1.812308],accel_mss,speed_ms,0,blend_radius_m)
  movel([0.241435, -1.332303, -2.582180, -0.797906, 1.570796, 1.812231],accel_mss,speed_ms,0,blend_radius_m)
  movel([0.241364, -1.332291, -2.582188, -0.797910, 1.570796, 1.812160],accel_mss,speed_ms,0,blend_radius_m)
  movel([0.235635, -1.330818, -2.583138, -0.798433, 1.570796, 1.806431],accel_mss,speed_ms,0,blend_radius_m)
  movel([0.229881, -1.329382, -2.584062, -0.798945, 1.570796, 1.800678],accel_mss,speed_ms,0,blend_radius_m)
  movel([0.229809, -1.329360, -2.584076, -0.798953, 1.570796, 1.800606],accel_mss,speed_ms,0,blend_radius_m)
  movel([0.229745, -1.329326, -2.584098, -0.798965, 1.570796, 1.800541],accel_mss,speed_ms,0,blend_radius_m)
  movel([0.229691, -1.329282, -2.584126, -0.798981, 1.570796, 1.800487],accel_mss,speed_ms,0,blend_radius_m)
  movel([0.229674, -1.329260, -2.584140, -0.798989, 1.570796, 1.800471],accel_mss,speed_ms,0,blend_radius_m)
  movel([0.229674, -1.329230, -2.584159, -0.798999, 1.570796, 1.800471],accel_mss,speed_ms,0,blend_radius_m)
  movel([0.229683, -1.329197, -2.584181, -0.799011, 1.570796, 1.800479],accel_mss,speed_ms,0,blend_radius_m)
  movel([0.231360, -1.325661, -2.586443, -0.800285, 1.570796, 1.802156],accel_mss,speed_ms,0,blend_radius_m)
  movel([0.233035, -1.322137, -2.588681, -0.801571, 1.570796, 1.803831],accel_mss,speed_ms,0,blend_radius_m)
  movel([0.233066, -1.322081, -2.588716, -0.801592, 1.570796, 1.803862],accel_mss,speed_ms,0,blend_radius_m)
  movel([0.233110, -1.322024, -2.588752, -0.801613, 1.570796, 1.803906],accel_mss,speed_ms,0,blend_radius_m)
  movel([0.233159, -1.321974, -2.588784, -0.801631, 1.570796, 1.803955],accel_mss,speed_ms,0,blend_radius_m)
  movel([0.233188, -1.321957, -2.588795, -0.801638, 1.570796, 1.803984],accel_mss,speed_ms,0,blend_radius_m)
  movel([0.233215, -1.321956, -2.588795, -0.801638, 1.570796, 1.804011],accel_mss,speed_ms,0,blend_radius_m)
  movel([0.234264, -1.322394, -2.588518, -0.801477, 1.570796, 1.805060],accel_mss,speed_ms,0,blend_radius_m)
  movel([0.235432, -1.322895, -2.588201, -0.801293, 1.570796, 1.806228],accel_mss,speed_ms,0,blend_radius_m)
  movel([0.236807, -1.323503, -2.587815, -0.801071, 1.570796, 1.807603],accel_mss,speed_ms,0,blend_radius_m)
  movel([0.240394, -1.325077, -2.586815, -0.800497, 1.570796, 1.811190],accel_mss,speed_ms,0,blend_radius_m)
  movel([0.240464, -1.324984, -2.586874, -0.800531, 1.570796, 1.811261],accel_mss,speed_ms,0,blend_radius_m)
  movel([0.240519, -1.324887, -2.586936, -0.800566, 1.570796, 1.811315],accel_mss,speed_ms,0,blend_radius_m)
  movel([0.243670, -1.317933, -2.591329, -0.803127, 1.570796, 1.814466],accel_mss,speed_ms,0,blend_radius_m)
  movel([0.243670, -1.317868, -2.591370, -0.803151, 1.570796, 1.814466],accel_mss,speed_ms,0,blend_radius_m)
  movel([0.243650, -1.317842, -2.591386, -0.803161, 1.570796, 1.814446],accel_mss,speed_ms,0,blend_radius_m)
  movel([0.243610, -1.317844, -2.591385, -0.803160, 1.570796, 1.814407],accel_mss,speed_ms,0,blend_radius_m)
  movel([0.240415, -1.318956, -2.590687, -0.802746, 1.570796, 1.811211],accel_mss,speed_ms,0,blend_radius_m)
  movel([0.236381, -1.320430, -2.589759, -0.802200, 1.570796, 1.807177],accel_mss,speed_ms,0,blend_radius_m)
  movel([0.234677, -1.321046, -2.589370, -0.801973, 1.570796, 1.805473],accel_mss,speed_ms,0,blend_radius_m)
  movel([0.233161, -1.321590, -2.589027, -0.801773, 1.570796, 1.803957],accel_mss,speed_ms,0,blend_radius_m)
  movel([0.233128, -1.321594, -2.589024, -0.801771, 1.570796, 1.803924],accel_mss,speed_ms,0,blend_radius_m)
  movel([0.233104, -1.321582, -2.589032, -0.801775, 1.570796, 1.803900],accel_mss,speed_ms,0,blend_radius_m)
  movel([0.233092, -1.321561, -2.589045, -0.801783, 1.570796, 1.803889],accel_mss,speed_ms,0,blend_radius_m)
  movel([0.233089, -1.321534, -2.589062, -0.801793, 1.570796, 1.803886],accel_mss,speed_ms,0,blend_radius_m)
  movel([0.233099, -1.321505, -2.589080, -0.801804, 1.570796, 1.803895],accel_mss,speed_ms,0,blend_radius_m)
  movel([0.234740, -1.318110, -2.591218, -0.803061, 1.570796, 1.805536],accel_mss,speed_ms,0,blend_radius_m)
  movel([0.236366, -1.314748, -2.593320, -0.804321, 1.570796, 1.807163],accel_mss,speed_ms,0,blend_radius_m)
  movel([0.236406, -1.314681, -2.593362, -0.804347, 1.570796, 1.807202],accel_mss,speed_ms,0,blend_radius_m)
  movel([0.236450, -1.314614, -2.593403, -0.804372, 1.570796, 1.807246],accel_mss,speed_ms,0,blend_radius_m)
  movel([0.236506, -1.314550, -2.593443, -0.804396, 1.570796, 1.807302],accel_mss,speed_ms,0,blend_radius_m)
  movel([0.236518, -1.314539, -2.593450, -0.804400, 1.570796, 1.807315],accel_mss,speed_ms,0,blend_radius_m)
  movel([0.236535, -1.314531, -2.593455, -0.804403, 1.570796, 1.807331],accel_mss,speed_ms,0,blend_radius_m)
  movel([0.239167, -1.313519, -2.594084, -0.804785, 1.570796, 1.809963],accel_mss,speed_ms,0,blend_radius_m)
  movel([0.242080, -1.312406, -2.594775, -0.805207, 1.570796, 1.812877],accel_mss,speed_ms,0,blend_radius_m)
  movel([0.245538, -1.311098, -2.595585, -0.805706, 1.570796, 1.816334],accel_mss,speed_ms,0,blend_radius_m)
  movel([0.254573, -1.307721, -2.597666, -0.807002, 1.570796, 1.825369],accel_mss,speed_ms,0,blend_radius_m)
  movel([0.256712, -1.309975, -2.596279, -0.806135, 1.570796, 1.827508],accel_mss,speed_ms,0,blend_radius_m)
  movel([0.258834, -1.312234, -2.594882, -0.805273, 1.570796, 1.829630],accel_mss,speed_ms,0,blend_radius_m)
  movel([0.258249, -1.313344, -2.594193, -0.804852, 1.570796, 1.829045],accel_mss,speed_ms,0,blend_radius_m)
  movel([0.257718, -1.314515, -2.593465, -0.804409, 1.570796, 1.828515],accel_mss,speed_ms,0,blend_radius_m)
  movel([0.257784, -1.314560, -2.593437, -0.804392, 1.570796, 1.828581],accel_mss,speed_ms,0,blend_radius_m)
  movel([0.257869, -1.314581, -2.593424, -0.804384, 1.570796, 1.828666],accel_mss,speed_ms,0,blend_radius_m)
  movel([0.260957, -1.314813, -2.593280, -0.804297, 1.570796, 1.831753],accel_mss,speed_ms,0,blend_radius_m)
  movel([0.266885, -1.315232, -2.593018, -0.804139, 1.570796, 1.837682],accel_mss,speed_ms,0,blend_radius_m)
  movel([0.268895, -1.315390, -2.592920, -0.804079, 1.570796, 1.839691],accel_mss,speed_ms,0,blend_radius_m)
  movel([0.270215, -1.315507, -2.592847, -0.804035, 1.570796, 1.841011],accel_mss,speed_ms,0,blend_radius_m)
  movel([0.271527, -1.315638, -2.592765, -0.803986, 1.570796, 1.842324],accel_mss,speed_ms,0,blend_radius_m)
  movel([0.272559, -1.315758, -2.592690, -0.803941, 1.570796, 1.843355],accel_mss,speed_ms,0,blend_radius_m)
  movel([0.273581, -1.315892, -2.592606, -0.803891, 1.570796, 1.844378],accel_mss,speed_ms,0,blend_radius_m)
  movel([0.274595, -1.316045, -2.592511, -0.803833, 1.570796, 1.845392],accel_mss,speed_ms,0,blend_radius_m)
  movel([0.275600, -1.316212, -2.592406, -0.803770, 1.570796, 1.846396],accel_mss,speed_ms,0,blend_radius_m)
  movel([0.276477, -1.316379, -2.592302, -0.803708, 1.570796, 1.847273],accel_mss,speed_ms,0,blend_radius_m)
  movel([0.277342, -1.316562, -2.592188, -0.803639, 1.570796, 1.848138],accel_mss,speed_ms,0,blend_radius_m)
  movel([0.278192, -1.316767, -2.592059, -0.803563, 1.570796, 1.848989],accel_mss,speed_ms,0,blend_radius_m)
  movel([0.279033, -1.316988, -2.591921, -0.803480, 1.570796, 1.849829],accel_mss,speed_ms,0,blend_radius_m)
  movel([0.279859, -1.317228, -2.591771, -0.803390, 1.570796, 1.850656],accel_mss,speed_ms,0,blend_radius_m)
  movel([0.280672, -1.317487, -2.591608, -0.803293, 1.570796, 1.851469],accel_mss,speed_ms,0,blend_radius_m)
  movel([0.281147, -1.317656, -2.591502, -0.803230, 1.570796, 1.851944],accel_mss,speed_ms,0,blend_radius_m)
  movel([0.281608, -1.317839, -2.591388, -0.803162, 1.570796, 1.852404],accel_mss,speed_ms,0,blend_radius_m)
  movel([0.282056, -1.318038, -2.591263, -0.803088, 1.570796, 1.852853],accel_mss,speed_ms,0,blend_radius_m)
  movel([0.282492, -1.318253, -2.591128, -0.803008, 1.570796, 1.853288],accel_mss,speed_ms,0,blend_radius_m)
  movel([0.282917, -1.318482, -2.590985, -0.802923, 1.570796, 1.853713],accel_mss,speed_ms,0,blend_radius_m)
  movel([0.283326, -1.318727, -2.590831, -0.802832, 1.570796, 1.854122],accel_mss,speed_ms,0,blend_radius_m)
  movel([0.283723, -1.318987, -2.590667, -0.802735, 1.570796, 1.854519],accel_mss,speed_ms,0,blend_radius_m)
  movel([0.284104, -1.319260, -2.590496, -0.802634, 1.570796, 1.854900],accel_mss,speed_ms,0,blend_radius_m)
  movel([0.284411, -1.319503, -2.590342, -0.802543, 1.570796, 1.855208],accel_mss,speed_ms,0,blend_radius_m)
  movel([0.284702, -1.319761, -2.590180, -0.802448, 1.570796, 1.855498],accel_mss,speed_ms,0,blend_radius_m)
  movel([0.284978, -1.320035, -2.590008, -0.802346, 1.570796, 1.855774],accel_mss,speed_ms,0,blend_radius_m)
  movel([0.285237, -1.320320, -2.589828, -0.802241, 1.570796, 1.856034],accel_mss,speed_ms,0,blend_radius_m)
  movel([0.285480, -1.320622, -2.589638, -0.802130, 1.570796, 1.856276],accel_mss,speed_ms,0,blend_radius_m)
  movel([0.285707, -1.320935, -2.589440, -0.802014, 1.570796, 1.856503],accel_mss,speed_ms,0,blend_radius_m)
  movel([0.285918, -1.321259, -2.589235, -0.801894, 1.570796, 1.856714],accel_mss,speed_ms,0,blend_radius_m)
  movel([0.286109, -1.321601, -2.589020, -0.801768, 1.570796, 1.856905],accel_mss,speed_ms,0,blend_radius_m)
  movel([0.286274, -1.321932, -2.588810, -0.801647, 1.570796, 1.857070],accel_mss,speed_ms,0,blend_radius_m)
  movel([0.286415, -1.322275, -2.588593, -0.801521, 1.570796, 1.857212],accel_mss,speed_ms,0,blend_radius_m)
  movel([0.286541, -1.322632, -2.588367, -0.801390, 1.570796, 1.857337],accel_mss,speed_ms,0,blend_radius_m)
  movel([0.286643, -1.323002, -2.588133, -0.801254, 1.570796, 1.857439],accel_mss,speed_ms,0,blend_radius_m)
  movel([0.286727, -1.323381, -2.587893, -0.801116, 1.570796, 1.857523],accel_mss,speed_ms,0,blend_radius_m)
  movel([0.286788, -1.323772, -2.587644, -0.800973, 1.570796, 1.857585],accel_mss,speed_ms,0,blend_radius_m)
  movel([0.286832, -1.324173, -2.587390, -0.800826, 1.570796, 1.857629],accel_mss,speed_ms,0,blend_radius_m)
  movel([0.286854, -1.324580, -2.587131, -0.800678, 1.570796, 1.857651],accel_mss,speed_ms,0,blend_radius_m)
  movel([0.286852, -1.324838, -2.586967, -0.800584, 1.570796, 1.857649],accel_mss,speed_ms,0,blend_radius_m)
  movel([0.286837, -1.325102, -2.586799, -0.800488, 1.570796, 1.857633],accel_mss,speed_ms,0,blend_radius_m)
  movel([0.286805, -1.325371, -2.586628, -0.800390, 1.570796, 1.857601],accel_mss,speed_ms,0,blend_radius_m)
  movel([0.286757, -1.325644, -2.586454, -0.800291, 1.570796, 1.857553],accel_mss,speed_ms,0,blend_radius_m)
  movel([0.286649, -1.326155, -2.586128, -0.800106, 1.570796, 1.857445],accel_mss,speed_ms,0,blend_radius_m)
  movel([0.286529, -1.326664, -2.585803, -0.799922, 1.570796, 1.857325],accel_mss,speed_ms,0,blend_radius_m)
  movel([0.286393, -1.327178, -2.585475, -0.799737, 1.570796, 1.857189],accel_mss,speed_ms,0,blend_radius_m)
  movel([0.286238, -1.327707, -2.585136, -0.799546, 1.570796, 1.857034],accel_mss,speed_ms,0,blend_radius_m)
  movel([0.286068, -1.328236, -2.584797, -0.799356, 1.570796, 1.856865],accel_mss,speed_ms,0,blend_radius_m)
  movel([0.285886, -1.328769, -2.584456, -0.799165, 1.570796, 1.856682],accel_mss,speed_ms,0,blend_radius_m)
  movel([0.285764, -1.329087, -2.584251, -0.799051, 1.570796, 1.856561],accel_mss,speed_ms,0,blend_radius_m)
  movel([0.285633, -1.329407, -2.584046, -0.798936, 1.570796, 1.856429],accel_mss,speed_ms,0,blend_radius_m)
  movel([0.285488, -1.329724, -2.583842, -0.798823, 1.570796, 1.856284],accel_mss,speed_ms,0,blend_radius_m)
  movel([0.285332, -1.330045, -2.583636, -0.798708, 1.570796, 1.856129],accel_mss,speed_ms,0,blend_radius_m)
  movel([0.285175, -1.330347, -2.583442, -0.798600, 1.570796, 1.855971],accel_mss,speed_ms,0,blend_radius_m)
  movel([0.285014, -1.330647, -2.583248, -0.798493, 1.570796, 1.855810],accel_mss,speed_ms,0,blend_radius_m)
  movel([0.284916, -1.330810, -2.583143, -0.798436, 1.570796, 1.855712],accel_mss,speed_ms,0,blend_radius_m)
  movel([0.284805, -1.330970, -2.583040, -0.798379, 1.570796, 1.855601],accel_mss,speed_ms,0,blend_radius_m)
  movel([0.284743, -1.331047, -2.582990, -0.798351, 1.570796, 1.855539],accel_mss,speed_ms,0,blend_radius_m)
  movel([0.284675, -1.331121, -2.582943, -0.798325, 1.570796, 1.855471],accel_mss,speed_ms,0,blend_radius_m)
  movel([0.284598, -1.331191, -2.582898, -0.798300, 1.570796, 1.855394],accel_mss,speed_ms,0,blend_radius_m)
  movel([0.284458, -1.331305, -2.582825, -0.798260, 1.570796, 1.855254],accel_mss,speed_ms,0,blend_radius_m)
  movel([0.284314, -1.331407, -2.582759, -0.798223, 1.570796, 1.855110],accel_mss,speed_ms,0,blend_radius_m)
  movel([0.283941, -1.331688, -2.582578, -0.798124, 1.570796, 1.854737],accel_mss,speed_ms,0,blend_radius_m)
  movel([0.283919, -1.331727, -2.582552, -0.798110, 1.570796, 1.854716],accel_mss,speed_ms,0,blend_radius_m)
  movel([0.283920, -1.331764, -2.582528, -0.798097, 1.570796, 1.854716],accel_mss,speed_ms,0,blend_radius_m)
  movel([0.283970, -1.331844, -2.582476, -0.798068, 1.570796, 1.854766],accel_mss,speed_ms,0,blend_radius_m)
  movel([0.284002, -1.331881, -2.582452, -0.798055, 1.570796, 1.854798],accel_mss,speed_ms,0,blend_radius_m)
  movel([0.284021, -1.331927, -2.582423, -0.798039, 1.570796, 1.854818],accel_mss,speed_ms,0,blend_radius_m)
  movel([0.284026, -1.331981, -2.582388, -0.798020, 1.570796, 1.854823],accel_mss,speed_ms,0,blend_radius_m)
  movel([0.284018, -1.332040, -2.582350, -0.797999, 1.570796, 1.854814],accel_mss,speed_ms,0,blend_radius_m)
  movel([0.283876, -1.332578, -2.582003, -0.797809, 1.570796, 1.854672],accel_mss,speed_ms,0,blend_radius_m)
  movel([0.283729, -1.333116, -2.581655, -0.797619, 1.570796, 1.854525],accel_mss,speed_ms,0,blend_radius_m)
  movel([0.283482, -1.333990, -2.581088, -0.797311, 1.570796, 1.854278],accel_mss,speed_ms,0,blend_radius_m)
  movel([0.283223, -1.334864, -2.580521, -0.797004, 1.570796, 1.854019],accel_mss,speed_ms,0,blend_radius_m)
  movel([0.282103, -1.338565, -2.578108, -0.795716, 1.570796, 1.852899],accel_mss,speed_ms,0,blend_radius_m)
  movel([0.280125, -1.345098, -2.573803, -0.793488, 1.570796, 1.850921],accel_mss,speed_ms,0,blend_radius_m)
  movel([0.282569, -1.344743, -2.574038, -0.793608, 1.570796, 1.853365],accel_mss,speed_ms,0,blend_radius_m)
  movel([0.285010, -1.344392, -2.574271, -0.793726, 1.570796, 1.855806],accel_mss,speed_ms,0,blend_radius_m)
  movel([0.286729, -1.340036, -2.577143, -0.795210, 1.570796, 1.857525],accel_mss,speed_ms,0,blend_radius_m)
  movel([0.287401, -1.338334, -2.578259, -0.795796, 1.570796, 1.858198],accel_mss,speed_ms,0,blend_radius_m)
  movel([0.287994, -1.336838, -2.579236, -0.796315, 1.570796, 1.858791],accel_mss,speed_ms,0,blend_radius_m)
  movel([0.288505, -1.335558, -2.580070, -0.796761, 1.570796, 1.859301],accel_mss,speed_ms,0,blend_radius_m)
  movel([0.288608, -1.335300, -2.580238, -0.796851, 1.570796, 1.859405],accel_mss,speed_ms,0,blend_radius_m)
  movel([0.288648, -1.335219, -2.580290, -0.796880, 1.570796, 1.859444],accel_mss,speed_ms,0,blend_radius_m)
  movel([0.288693, -1.335143, -2.580340, -0.796906, 1.570796, 1.859489],accel_mss,speed_ms,0,blend_radius_m)
  movel([0.288753, -1.335057, -2.580396, -0.796936, 1.570796, 1.859549],accel_mss,speed_ms,0,blend_radius_m)
  movel([0.288819, -1.334975, -2.580449, -0.796965, 1.570796, 1.859615],accel_mss,speed_ms,0,blend_radius_m)
  movel([0.288894, -1.334894, -2.580501, -0.796993, 1.570796, 1.859690],accel_mss,speed_ms,0,blend_radius_m)
  movel([0.288973, -1.334818, -2.580551, -0.797020, 1.570796, 1.859769],accel_mss,speed_ms,0,blend_radius_m)
  movel([0.289051, -1.334750, -2.580595, -0.797044, 1.570796, 1.859847],accel_mss,speed_ms,0,blend_radius_m)
  movel([0.289131, -1.334692, -2.580633, -0.797064, 1.570796, 1.859927],accel_mss,speed_ms,0,blend_radius_m)
  movel([0.289240, -1.334625, -2.580676, -0.797088, 1.570796, 1.860037],accel_mss,speed_ms,0,blend_radius_m)
  movel([0.289355, -1.334571, -2.580711, -0.797107, 1.570796, 1.860151],accel_mss,speed_ms,0,blend_radius_m)
  movel([0.289466, -1.334536, -2.580734, -0.797119, 1.570796, 1.860262],accel_mss,speed_ms,0,blend_radius_m)
  movel([0.289621, -1.334499, -2.580758, -0.797132, 1.570796, 1.860417],accel_mss,speed_ms,0,blend_radius_m)
  movel([0.289775, -1.334470, -2.580777, -0.797142, 1.570796, 1.860572],accel_mss,speed_ms,0,blend_radius_m)
  movel([0.289924, -1.334453, -2.580788, -0.797148, 1.570796, 1.860720],accel_mss,speed_ms,0,blend_radius_m)
  movel([0.290333, -1.334418, -2.580810, -0.797160, 1.570796, 1.861130],accel_mss,speed_ms,0,blend_radius_m)
  movel([0.290736, -1.334398, -2.580823, -0.797167, 1.570796, 1.861532],accel_mss,speed_ms,0,blend_radius_m)
  movel([0.292944, -1.334330, -2.580868, -0.797191, 1.570796, 1.863740],accel_mss,speed_ms,0,blend_radius_m)
  movel([0.294287, -1.334295, -2.580890, -0.797204, 1.570796, 1.865083],accel_mss,speed_ms,0,blend_radius_m)
  movel([0.295478, -1.334270, -2.580907, -0.797213, 1.570796, 1.866275],accel_mss,speed_ms,0,blend_radius_m)
  movel([0.296484, -1.334252, -2.580918, -0.797219, 1.570796, 1.867280],accel_mss,speed_ms,0,blend_radius_m)
  movel([0.296752, -1.334256, -2.580916, -0.797217, 1.570796, 1.867549],accel_mss,speed_ms,0,blend_radius_m)
  movel([0.296861, -1.334265, -2.580910, -0.797214, 1.570796, 1.867658],accel_mss,speed_ms,0,blend_radius_m)
  movel([0.296966, -1.334282, -2.580899, -0.797208, 1.570796, 1.867762],accel_mss,speed_ms,0,blend_radius_m)
  movel([0.297062, -1.334309, -2.580881, -0.797199, 1.570796, 1.867858],accel_mss,speed_ms,0,blend_radius_m)
  movel([0.297138, -1.334341, -2.580860, -0.797187, 1.570796, 1.867934],accel_mss,speed_ms,0,blend_radius_m)
  movel([0.297202, -1.334386, -2.580831, -0.797172, 1.570796, 1.867999],accel_mss,speed_ms,0,blend_radius_m)
  movel([0.297254, -1.334442, -2.580795, -0.797152, 1.570796, 1.868050],accel_mss,speed_ms,0,blend_radius_m)
  movel([0.297294, -1.334503, -2.580755, -0.797130, 1.570796, 1.868090],accel_mss,speed_ms,0,blend_radius_m)
  movel([0.297317, -1.334574, -2.580709, -0.797106, 1.570796, 1.868113],accel_mss,speed_ms,0,blend_radius_m)
  movel([0.297328, -1.334651, -2.580660, -0.797079, 1.570796, 1.868124],accel_mss,speed_ms,0,blend_radius_m)
  movel([0.297325, -1.334743, -2.580600, -0.797046, 1.570796, 1.868121],accel_mss,speed_ms,0,blend_radius_m)
  movel([0.297312, -1.334836, -2.580539, -0.797014, 1.570796, 1.868108],accel_mss,speed_ms,0,blend_radius_m)
  movel([0.297286, -1.334934, -2.580476, -0.796980, 1.570796, 1.868082],accel_mss,speed_ms,0,blend_radius_m)
  movel([0.297243, -1.335120, -2.580355, -0.796914, 1.570796, 1.868039],accel_mss,speed_ms,0,blend_radius_m)
  movel([0.297264, -1.335218, -2.580291, -0.796880, 1.570796, 1.868060],accel_mss,speed_ms,0,blend_radius_m)
  movel([0.297355, -1.335269, -2.580258, -0.796862, 1.570796, 1.868151],accel_mss,speed_ms,0,blend_radius_m)
  movel([0.297561, -1.335290, -2.580244, -0.796855, 1.570796, 1.868357],accel_mss,speed_ms,0,blend_radius_m)
  movel([0.297762, -1.335295, -2.580241, -0.796853, 1.570796, 1.868558],accel_mss,speed_ms,0,blend_radius_m)
  movel([0.298076, -1.335302, -2.580236, -0.796851, 1.570796, 1.868872],accel_mss,speed_ms,0,blend_radius_m)
  movel([0.298427, -1.335315, -2.580228, -0.796846, 1.570796, 1.869224],accel_mss,speed_ms,0,blend_radius_m)
  movel([0.298770, -1.335323, -2.580222, -0.796843, 1.570796, 1.869566],accel_mss,speed_ms,0,blend_radius_m)
  movel([0.299314, -1.335349, -2.580206, -0.796834, 1.570796, 1.870111],accel_mss,speed_ms,0,blend_radius_m)
  movel([0.299852, -1.335388, -2.580181, -0.796821, 1.570796, 1.870649],accel_mss,speed_ms,0,blend_radius_m)
  movel([0.300380, -1.335443, -2.580144, -0.796801, 1.570796, 1.871176],accel_mss,speed_ms,0,blend_radius_m)
  movel([0.300900, -1.335514, -2.580098, -0.796776, 1.570796, 1.871697],accel_mss,speed_ms,0,blend_radius_m)
  movel([0.301411, -1.335600, -2.580042, -0.796746, 1.570796, 1.872207],accel_mss,speed_ms,0,blend_radius_m)
  movel([0.301911, -1.335702, -2.579976, -0.796711, 1.570796, 1.872708],accel_mss,speed_ms,0,blend_radius_m)
  movel([0.302405, -1.335818, -2.579901, -0.796670, 1.570796, 1.873201],accel_mss,speed_ms,0,blend_radius_m)
  movel([0.302886, -1.335949, -2.579815, -0.796624, 1.570796, 1.873682],accel_mss,speed_ms,0,blend_radius_m)
  movel([0.303443, -1.336123, -2.579702, -0.796564, 1.570796, 1.874240],accel_mss,speed_ms,0,blend_radius_m)
  movel([0.303985, -1.336314, -2.579577, -0.796497, 1.570796, 1.874782],accel_mss,speed_ms,0,blend_radius_m)
  movel([0.304516, -1.336526, -2.579439, -0.796423, 1.570796, 1.875312],accel_mss,speed_ms,0,blend_radius_m)
  movel([0.305031, -1.336753, -2.579291, -0.796344, 1.570796, 1.875828],accel_mss,speed_ms,0,blend_radius_m)
  movel([0.305534, -1.336999, -2.579131, -0.796259, 1.570796, 1.876330],accel_mss,speed_ms,0,blend_radius_m)
  movel([0.306018, -1.337262, -2.578959, -0.796168, 1.570796, 1.876814],accel_mss,speed_ms,0,blend_radius_m)
  movel([0.306489, -1.337544, -2.578775, -0.796070, 1.570796, 1.877285],accel_mss,speed_ms,0,blend_radius_m)
  movel([0.306951, -1.337842, -2.578580, -0.795966, 1.570796, 1.877747],accel_mss,speed_ms,0,blend_radius_m)
  movel([0.307394, -1.338161, -2.578372, -0.795856, 1.570796, 1.878191],accel_mss,speed_ms,0,blend_radius_m)
  movel([0.307824, -1.338494, -2.578154, -0.795741, 1.570796, 1.878620],accel_mss,speed_ms,0,blend_radius_m)
  movel([0.308235, -1.338844, -2.577925, -0.795620, 1.570796, 1.879031],accel_mss,speed_ms,0,blend_radius_m)
  movel([0.308631, -1.339210, -2.577685, -0.795494, 1.570796, 1.879427],accel_mss,speed_ms,0,blend_radius_m)
  movel([0.309007, -1.339592, -2.577435, -0.795362, 1.570796, 1.879803],accel_mss,speed_ms,0,blend_radius_m)
  movel([0.309367, -1.339987, -2.577175, -0.795226, 1.570796, 1.880163],accel_mss,speed_ms,0,blend_radius_m)
  movel([0.309705, -1.340396, -2.576907, -0.795086, 1.570796, 1.880501],accel_mss,speed_ms,0,blend_radius_m)
  movel([0.310025, -1.340817, -2.576630, -0.794942, 1.570796, 1.880821],accel_mss,speed_ms,0,blend_radius_m)
  movel([0.310324, -1.341255, -2.576342, -0.794792, 1.570796, 1.881120],accel_mss,speed_ms,0,blend_radius_m)
  movel([0.310607, -1.341704, -2.576046, -0.794639, 1.570796, 1.881404],accel_mss,speed_ms,0,blend_radius_m)
  movel([0.310869, -1.342169, -2.575740, -0.794480, 1.570796, 1.881665],accel_mss,speed_ms,0,blend_radius_m)
  movel([0.311114, -1.342645, -2.575426, -0.794318, 1.570796, 1.881911],accel_mss,speed_ms,0,blend_radius_m)
  movel([0.311336, -1.343134, -2.575103, -0.794152, 1.570796, 1.882132],accel_mss,speed_ms,0,blend_radius_m)
  movel([0.311538, -1.343625, -2.574778, -0.793986, 1.570796, 1.882334],accel_mss,speed_ms,0,blend_radius_m)
  movel([0.311719, -1.344130, -2.574444, -0.793815, 1.570796, 1.882515],accel_mss,speed_ms,0,blend_radius_m)
  movel([0.311882, -1.344643, -2.574104, -0.793642, 1.570796, 1.882678],accel_mss,speed_ms,0,blend_radius_m)
  movel([0.312027, -1.345166, -2.573757, -0.793465, 1.570796, 1.882824],accel_mss,speed_ms,0,blend_radius_m)
  movel([0.312152, -1.345701, -2.573402, -0.793286, 1.570796, 1.882949],accel_mss,speed_ms,0,blend_radius_m)
  movel([0.312266, -1.346275, -2.573021, -0.793093, 1.570796, 1.883063],accel_mss,speed_ms,0,blend_radius_m)
  movel([0.312363, -1.346857, -2.572633, -0.792898, 1.570796, 1.883159],accel_mss,speed_ms,0,blend_radius_m)
  movel([0.312445, -1.347447, -2.572240, -0.792701, 1.570796, 1.883242],accel_mss,speed_ms,0,blend_radius_m)
  movel([0.312508, -1.348046, -2.571841, -0.792502, 1.570796, 1.883304],accel_mss,speed_ms,0,blend_radius_m)
  movel([0.312554, -1.348650, -2.571438, -0.792301, 1.570796, 1.883351],accel_mss,speed_ms,0,blend_radius_m)
  movel([0.312581, -1.349249, -2.571037, -0.792103, 1.570796, 1.883377],accel_mss,speed_ms,0,blend_radius_m)
  movel([0.312592, -1.349851, -2.570634, -0.791904, 1.570796, 1.883389],accel_mss,speed_ms,0,blend_radius_m)
  movel([0.312587, -1.350462, -2.570225, -0.791702, 1.570796, 1.883383],accel_mss,speed_ms,0,blend_radius_m)
  movel([0.312566, -1.351075, -2.569813, -0.791501, 1.570796, 1.883363],accel_mss,speed_ms,0,blend_radius_m)
  movel([0.312526, -1.351697, -2.569396, -0.791297, 1.570796, 1.883322],accel_mss,speed_ms,0,blend_radius_m)
  movel([0.312484, -1.352163, -2.569082, -0.791144, 1.570796, 1.883281],accel_mss,speed_ms,0,blend_radius_m)
  movel([0.312427, -1.352635, -2.568764, -0.790990, 1.570796, 1.883223],accel_mss,speed_ms,0,blend_radius_m)
  movel([0.312354, -1.353110, -2.568444, -0.790835, 1.570796, 1.883150],accel_mss,speed_ms,0,blend_radius_m)
  movel([0.312268, -1.353588, -2.568121, -0.790679, 1.570796, 1.883064],accel_mss,speed_ms,0,blend_radius_m)
  movel([0.312170, -1.354070, -2.567796, -0.790523, 1.570796, 1.882966],accel_mss,speed_ms,0,blend_radius_m)
  movel([0.312054, -1.354553, -2.567470, -0.790366, 1.570796, 1.882851],accel_mss,speed_ms,0,blend_radius_m)
  movel([0.311928, -1.355174, -2.567050, -0.790166, 1.570796, 1.882724],accel_mss,speed_ms,0,blend_radius_m)
  movel([0.311926, -1.355257, -2.566993, -0.790139, 1.570796, 1.882722],accel_mss,speed_ms,0,blend_radius_m)
  movel([0.311951, -1.355326, -2.566947, -0.790116, 1.570796, 1.882748],accel_mss,speed_ms,0,blend_radius_m)
  movel([0.312001, -1.355379, -2.566910, -0.790099, 1.570796, 1.882797],accel_mss,speed_ms,0,blend_radius_m)
  movel([0.312125, -1.355434, -2.566873, -0.790082, 1.570796, 1.882921],accel_mss,speed_ms,0,blend_radius_m)
  movel([0.312269, -1.355456, -2.566859, -0.790075, 1.570796, 1.883065],accel_mss,speed_ms,0,blend_radius_m)
  movel([0.313348, -1.355447, -2.566864, -0.790077, 1.570796, 1.884144],accel_mss,speed_ms,0,blend_radius_m)
  movel([0.314266, -1.355434, -2.566874, -0.790082, 1.570796, 1.885062],accel_mss,speed_ms,0,blend_radius_m)
  movel([0.314079, -1.355802, -2.566624, -0.789963, 1.570796, 1.884875],accel_mss,speed_ms,0,blend_radius_m)
  movel([0.313825, -1.356353, -2.566250, -0.789786, 1.570796, 1.884622],accel_mss,speed_ms,0,blend_radius_m)
  movel([0.312966, -1.358517, -2.564778, -0.789094, 1.570796, 1.883763],accel_mss,speed_ms,0,blend_radius_m)
  movel([0.312961, -1.358602, -2.564720, -0.789067, 1.570796, 1.883757],accel_mss,speed_ms,0,blend_radius_m)
  movel([0.312997, -1.358652, -2.564686, -0.789051, 1.570796, 1.883794],accel_mss,speed_ms,0,blend_radius_m)
  movel([0.314293, -1.359063, -2.564406, -0.788920, 1.570796, 1.885090],accel_mss,speed_ms,0,blend_radius_m)
  movel([0.314628, -1.359178, -2.564327, -0.788884, 1.570796, 1.885424],accel_mss,speed_ms,0,blend_radius_m)
  movel([0.314954, -1.359305, -2.564240, -0.788843, 1.570796, 1.885750],accel_mss,speed_ms,0,blend_radius_m)
  movel([0.315271, -1.359445, -2.564145, -0.788799, 1.570796, 1.886067],accel_mss,speed_ms,0,blend_radius_m)
  movel([0.315576, -1.359599, -2.564040, -0.788750, 1.570796, 1.886372],accel_mss,speed_ms,0,blend_radius_m)
  movel([0.315878, -1.359773, -2.563921, -0.788695, 1.570796, 1.886674],accel_mss,speed_ms,0,blend_radius_m)
  movel([0.316172, -1.359960, -2.563793, -0.788636, 1.570796, 1.886968],accel_mss,speed_ms,0,blend_radius_m)
  movel([0.316455, -1.360156, -2.563659, -0.788574, 1.570796, 1.887251],accel_mss,speed_ms,0,blend_radius_m)
  movel([0.316724, -1.360365, -2.563516, -0.788508, 1.570796, 1.887521],accel_mss,speed_ms,0,blend_radius_m)
  movel([0.316982, -1.360587, -2.563364, -0.788438, 1.570796, 1.887779],accel_mss,speed_ms,0,blend_radius_m)
  movel([0.317236, -1.360822, -2.563204, -0.788364, 1.570796, 1.888032],accel_mss,speed_ms,0,blend_radius_m)
  movel([0.317475, -1.361069, -2.563034, -0.788286, 1.570796, 1.888272],accel_mss,speed_ms,0,blend_radius_m)
  movel([0.317702, -1.361329, -2.562856, -0.788204, 1.570796, 1.888498],accel_mss,speed_ms,0,blend_radius_m)
  movel([0.317915, -1.361597, -2.562672, -0.788120, 1.570796, 1.888712],accel_mss,speed_ms,0,blend_radius_m)
  movel([0.318117, -1.361875, -2.562482, -0.788033, 1.570796, 1.888913],accel_mss,speed_ms,0,blend_radius_m)
  movel([0.318306, -1.362165, -2.562283, -0.787942, 1.570796, 1.889103],accel_mss,speed_ms,0,blend_radius_m)
  movel([0.318481, -1.362465, -2.562076, -0.787848, 1.570796, 1.889277],accel_mss,speed_ms,0,blend_radius_m)
  movel([0.318641, -1.362773, -2.561865, -0.787752, 1.570796, 1.889438],accel_mss,speed_ms,0,blend_radius_m)
  movel([0.318792, -1.363088, -2.561648, -0.787653, 1.570796, 1.889588],accel_mss,speed_ms,0,blend_radius_m)
  movel([0.318925, -1.363414, -2.561423, -0.787551, 1.570796, 1.889721],accel_mss,speed_ms,0,blend_radius_m)
  movel([0.319051, -1.363767, -2.561180, -0.787442, 1.570796, 1.889847],accel_mss,speed_ms,0,blend_radius_m)
  movel([0.319161, -1.364130, -2.560930, -0.787329, 1.570796, 1.889958],accel_mss,speed_ms,0,blend_radius_m)
  movel([0.319255, -1.364502, -2.560674, -0.787214, 1.570796, 1.890052],accel_mss,speed_ms,0,blend_radius_m)
  movel([0.319333, -1.364881, -2.560412, -0.787096, 1.570796, 1.890129],accel_mss,speed_ms,0,blend_radius_m)
  movel([0.319399, -1.365292, -2.560128, -0.786969, 1.570796, 1.890195],accel_mss,speed_ms,0,blend_radius_m)
  movel([0.319450, -1.365713, -2.559837, -0.786839, 1.570796, 1.890246],accel_mss,speed_ms,0,blend_radius_m)
  movel([0.319487, -1.366139, -2.559542, -0.786708, 1.570796, 1.890284],accel_mss,speed_ms,0,blend_radius_m)
  movel([0.319510, -1.366569, -2.559244, -0.786575, 1.570796, 1.890306],accel_mss,speed_ms,0,blend_radius_m)
  movel([0.319522, -1.367110, -2.558869, -0.786410, 1.570796, 1.890318],accel_mss,speed_ms,0,blend_radius_m)
  movel([0.319520, -1.367656, -2.558490, -0.786242, 1.570796, 1.890316],accel_mss,speed_ms,0,blend_radius_m)
  movel([0.319503, -1.368206, -2.558109, -0.786075, 1.570796, 1.890300],accel_mss,speed_ms,0,blend_radius_m)
  movel([0.319476, -1.368758, -2.557725, -0.785907, 1.570796, 1.890273],accel_mss,speed_ms,0,blend_radius_m)
  movel([0.319406, -1.369776, -2.557016, -0.785598, 1.570796, 1.890202],accel_mss,speed_ms,0,blend_radius_m)
  movel([0.319320, -1.370798, -2.556302, -0.785289, 1.570796, 1.890116],accel_mss,speed_ms,0,blend_radius_m)
  movel([0.319224, -1.371822, -2.555586, -0.784981, 1.570796, 1.890020],accel_mss,speed_ms,0,blend_radius_m)
  movel([0.319012, -1.374151, -2.553952, -0.784287, 1.570796, 1.889808],accel_mss,speed_ms,0,blend_radius_m)
  movel([0.318877, -1.376237, -2.552481, -0.783671, 1.570796, 1.889673],accel_mss,speed_ms,0,blend_radius_m)
  movel([0.318819, -1.378011, -2.551226, -0.783152, 1.570796, 1.889615],accel_mss,speed_ms,0,blend_radius_m)
  movel([0.318820, -1.378689, -2.550745, -0.782955, 1.570796, 1.889616],accel_mss,speed_ms,0,blend_radius_m)
  movel([0.318846, -1.379356, -2.550271, -0.782762, 1.570796, 1.889643],accel_mss,speed_ms,0,blend_radius_m)
  movel([0.318897, -1.380237, -2.549645, -0.782508, 1.570796, 1.889693],accel_mss,speed_ms,0,blend_radius_m)
  movel([0.319580, -1.379966, -2.549838, -0.782586, 1.570796, 1.890377],accel_mss,speed_ms,0,blend_radius_m)
  movel([0.319784, -1.379890, -2.549891, -0.782607, 1.570796, 1.890580],accel_mss,speed_ms,0,blend_radius_m)
  movel([0.319985, -1.379826, -2.549937, -0.782626, 1.570796, 1.890781],accel_mss,speed_ms,0,blend_radius_m)
  movel([0.320184, -1.379775, -2.549973, -0.782641, 1.570796, 1.890981],accel_mss,speed_ms,0,blend_radius_m)
  movel([0.320383, -1.379733, -2.550003, -0.782653, 1.570796, 1.891179],accel_mss,speed_ms,0,blend_radius_m)
  movel([0.320686, -1.379684, -2.550038, -0.782667, 1.570796, 1.891482],accel_mss,speed_ms,0,blend_radius_m)
  movel([0.320983, -1.379652, -2.550061, -0.782676, 1.570796, 1.891779],accel_mss,speed_ms,0,blend_radius_m)
  movel([0.321275, -1.379635, -2.550073, -0.782681, 1.570796, 1.892071],accel_mss,speed_ms,0,blend_radius_m)
  movel([0.321564, -1.379633, -2.550074, -0.782682, 1.570796, 1.892360],accel_mss,speed_ms,0,blend_radius_m)
  movel([0.321844, -1.379648, -2.550064, -0.782677, 1.570796, 1.892641],accel_mss,speed_ms,0,blend_radius_m)
  movel([0.322115, -1.379679, -2.550042, -0.782669, 1.570796, 1.892912],accel_mss,speed_ms,0,blend_radius_m)
  movel([0.322289, -1.379708, -2.550021, -0.782660, 1.570796, 1.893085],accel_mss,speed_ms,0,blend_radius_m)
  movel([0.322456, -1.379750, -2.549991, -0.782648, 1.570796, 1.893252],accel_mss,speed_ms,0,blend_radius_m)
  movel([0.322613, -1.379800, -2.549955, -0.782633, 1.570796, 1.893409],accel_mss,speed_ms,0,blend_radius_m)
  movel([0.322763, -1.379865, -2.549910, -0.782615, 1.570796, 1.893559],accel_mss,speed_ms,0,blend_radius_m)
  movel([0.322955, -1.379965, -2.549838, -0.782586, 1.570796, 1.893751],accel_mss,speed_ms,0,blend_radius_m)
  movel([0.323134, -1.380081, -2.549755, -0.782552, 1.570796, 1.893931],accel_mss,speed_ms,0,blend_radius_m)
  movel([0.323297, -1.380212, -2.549662, -0.782515, 1.570796, 1.894094],accel_mss,speed_ms,0,blend_radius_m)
  movel([0.323446, -1.380357, -2.549559, -0.782473, 1.570796, 1.894243],accel_mss,speed_ms,0,blend_radius_m)
  movel([0.323593, -1.380528, -2.549437, -0.782424, 1.570796, 1.894389],accel_mss,speed_ms,0,blend_radius_m)
  movel([0.323722, -1.380710, -2.549308, -0.782371, 1.570796, 1.894518],accel_mss,speed_ms,0,blend_radius_m)
  movel([0.323839, -1.380901, -2.549172, -0.782317, 1.570796, 1.894635],accel_mss,speed_ms,0,blend_radius_m)
  movel([0.323941, -1.381101, -2.549029, -0.782259, 1.570796, 1.894737],accel_mss,speed_ms,0,blend_radius_m)
  movel([0.324027, -1.381314, -2.548877, -0.782198, 1.570796, 1.894823],accel_mss,speed_ms,0,blend_radius_m)
  movel([0.324099, -1.381535, -2.548720, -0.782135, 1.570796, 1.894896],accel_mss,speed_ms,0,blend_radius_m)
  movel([0.324155, -1.381763, -2.548557, -0.782070, 1.570796, 1.894952],accel_mss,speed_ms,0,blend_radius_m)
  movel([0.324195, -1.381998, -2.548388, -0.782002, 1.570796, 1.894991],accel_mss,speed_ms,0,blend_radius_m)
  movel([0.324217, -1.382227, -2.548225, -0.781937, 1.570796, 1.895013],accel_mss,speed_ms,0,blend_radius_m)
  movel([0.324221, -1.382461, -2.548058, -0.781870, 1.570796, 1.895017],accel_mss,speed_ms,0,blend_radius_m)
  movel([0.324205, -1.382701, -2.547886, -0.781802, 1.570796, 1.895001],accel_mss,speed_ms,0,blend_radius_m)
  movel([0.324171, -1.382946, -2.547711, -0.781732, 1.570796, 1.894967],accel_mss,speed_ms,0,blend_radius_m)
  movel([0.324123, -1.383193, -2.547534, -0.781662, 1.570796, 1.894919],accel_mss,speed_ms,0,blend_radius_m)
  movel([0.324059, -1.383444, -2.547354, -0.781591, 1.570796, 1.894856],accel_mss,speed_ms,0,blend_radius_m)
  movel([0.323980, -1.383697, -2.547172, -0.781519, 1.570796, 1.894776],accel_mss,speed_ms,0,blend_radius_m)
  movel([0.323888, -1.383951, -2.546990, -0.781447, 1.570796, 1.894685],accel_mss,speed_ms,0,blend_radius_m)
  movel([0.323782, -1.384204, -2.546809, -0.781376, 1.570796, 1.894578],accel_mss,speed_ms,0,blend_radius_m)
  movel([0.323663, -1.384460, -2.546626, -0.781304, 1.570796, 1.894459],accel_mss,speed_ms,0,blend_radius_m)
  movel([0.323530, -1.384710, -2.546446, -0.781233, 1.570796, 1.894327],accel_mss,speed_ms,0,blend_radius_m)
  movel([0.323387, -1.384959, -2.546267, -0.781163, 1.570796, 1.894183],accel_mss,speed_ms,0,blend_radius_m)
  movel([0.323230, -1.385206, -2.546089, -0.781094, 1.570796, 1.894027],accel_mss,speed_ms,0,blend_radius_m)
  movel([0.323061, -1.385450, -2.545914, -0.781025, 1.570796, 1.893858],accel_mss,speed_ms,0,blend_radius_m)
  movel([0.322881, -1.385688, -2.545742, -0.780958, 1.570796, 1.893677],accel_mss,speed_ms,0,blend_radius_m)
  movel([0.322688, -1.385925, -2.545572, -0.780892, 1.570796, 1.893484],accel_mss,speed_ms,0,blend_radius_m)
  movel([0.322486, -1.386154, -2.545407, -0.780828, 1.570796, 1.893282],accel_mss,speed_ms,0,blend_radius_m)
  movel([0.322275, -1.386378, -2.545246, -0.780765, 1.570796, 1.893072],accel_mss,speed_ms,0,blend_radius_m)
  movel([0.322055, -1.386595, -2.545089, -0.780705, 1.570796, 1.892851],accel_mss,speed_ms,0,blend_radius_m)
  movel([0.321827, -1.386804, -2.544938, -0.780646, 1.570796, 1.892623],accel_mss,speed_ms,0,blend_radius_m)
  movel([0.321590, -1.387006, -2.544793, -0.780590, 1.570796, 1.892386],accel_mss,speed_ms,0,blend_radius_m)
  movel([0.321345, -1.387199, -2.544654, -0.780536, 1.570796, 1.892141],accel_mss,speed_ms,0,blend_radius_m)
  movel([0.321093, -1.387384, -2.544520, -0.780485, 1.570796, 1.891890],accel_mss,speed_ms,0,blend_radius_m)
  movel([0.320837, -1.387559, -2.544394, -0.780436, 1.570796, 1.891633],accel_mss,speed_ms,0,blend_radius_m)
  movel([0.320576, -1.387726, -2.544273, -0.780390, 1.570796, 1.891372],accel_mss,speed_ms,0,blend_radius_m)
  movel([0.320308, -1.387882, -2.544160, -0.780347, 1.570796, 1.891104],accel_mss,speed_ms,0,blend_radius_m)
  movel([0.320040, -1.388025, -2.544057, -0.780307, 1.570796, 1.890836],accel_mss,speed_ms,0,blend_radius_m)
  movel([0.319767, -1.388158, -2.543961, -0.780270, 1.570796, 1.890563],accel_mss,speed_ms,0,blend_radius_m)
  movel([0.319548, -1.388257, -2.543889, -0.780243, 1.570796, 1.890344],accel_mss,speed_ms,0,blend_radius_m)
  movel([0.319328, -1.388345, -2.543825, -0.780218, 1.570796, 1.890125],accel_mss,speed_ms,0,blend_radius_m)
  movel([0.319149, -1.388409, -2.543779, -0.780201, 1.570796, 1.889945],accel_mss,speed_ms,0,blend_radius_m)
  movel([0.318972, -1.388459, -2.543743, -0.780187, 1.570796, 1.889768],accel_mss,speed_ms,0,blend_radius_m)
  movel([0.318771, -1.388501, -2.543713, -0.780175, 1.570796, 1.889567],accel_mss,speed_ms,0,blend_radius_m)
  movel([0.318573, -1.388531, -2.543691, -0.780167, 1.570796, 1.889370],accel_mss,speed_ms,0,blend_radius_m)
  movel([0.318277, -1.388563, -2.543667, -0.780158, 1.570796, 1.889073],accel_mss,speed_ms,0,blend_radius_m)
  movel([0.317981, -1.388591, -2.543647, -0.780150, 1.570796, 1.888778],accel_mss,speed_ms,0,blend_radius_m)
  movel([0.317692, -1.388610, -2.543634, -0.780145, 1.570796, 1.888488],accel_mss,speed_ms,0,blend_radius_m)
  movel([0.317400, -1.388627, -2.543622, -0.780141, 1.570796, 1.888196],accel_mss,speed_ms,0,blend_radius_m)
  movel([0.317211, -1.388627, -2.543622, -0.780141, 1.570796, 1.888007],accel_mss,speed_ms,0,blend_radius_m)
  movel([0.317028, -1.388616, -2.543630, -0.780144, 1.570796, 1.887825],accel_mss,speed_ms,0,blend_radius_m)
  movel([0.316872, -1.388594, -2.543645, -0.780150, 1.570796, 1.887668],accel_mss,speed_ms,0,blend_radius_m)
  movel([0.316722, -1.388557, -2.543672, -0.780160, 1.570796, 1.887519],accel_mss,speed_ms,0,blend_radius_m)
  movel([0.316548, -1.388500, -2.543713, -0.780176, 1.570796, 1.887345],accel_mss,speed_ms,0,blend_radius_m)
  movel([0.316382, -1.388434, -2.543761, -0.780194, 1.570796, 1.887178],accel_mss,speed_ms,0,blend_radius_m)
  movel([0.316165, -1.388331, -2.543835, -0.780222, 1.570796, 1.886962],accel_mss,speed_ms,0,blend_radius_m)
  movel([0.315963, -1.388212, -2.543921, -0.780255, 1.570796, 1.886759],accel_mss,speed_ms,0,blend_radius_m)
  movel([0.315777, -1.388077, -2.544019, -0.780293, 1.570796, 1.886574],accel_mss,speed_ms,0,blend_radius_m)
  movel([0.315603, -1.387928, -2.544127, -0.780334, 1.570796, 1.886400],accel_mss,speed_ms,0,blend_radius_m)
  movel([0.315447, -1.387767, -2.544243, -0.780378, 1.570796, 1.886243],accel_mss,speed_ms,0,blend_radius_m)
  movel([0.315307, -1.387590, -2.544371, -0.780428, 1.570796, 1.886103],accel_mss,speed_ms,0,blend_radius_m)
  movel([0.315185, -1.387400, -2.544509, -0.780480, 1.570796, 1.885981],accel_mss,speed_ms,0,blend_radius_m)
  movel([0.315078, -1.387198, -2.544654, -0.780537, 1.570796, 1.885875],accel_mss,speed_ms,0,blend_radius_m)
  movel([0.314989, -1.386984, -2.544809, -0.780596, 1.570796, 1.885785],accel_mss,speed_ms,0,blend_radius_m)
  movel([0.314920, -1.386758, -2.544972, -0.780659, 1.570796, 1.885716],accel_mss,speed_ms,0,blend_radius_m)
  movel([0.314867, -1.386523, -2.545141, -0.780725, 1.570796, 1.885663],accel_mss,speed_ms,0,blend_radius_m)
  movel([0.314832, -1.386281, -2.545316, -0.780792, 1.570796, 1.885629],accel_mss,speed_ms,0,blend_radius_m)
  movel([0.314817, -1.386028, -2.545498, -0.780863, 1.570796, 1.885613],accel_mss,speed_ms,0,blend_radius_m)
  movel([0.314820, -1.385770, -2.545684, -0.780935, 1.570796, 1.885616],accel_mss,speed_ms,0,blend_radius_m)
  movel([0.314840, -1.385505, -2.545874, -0.781010, 1.570796, 1.885636],accel_mss,speed_ms,0,blend_radius_m)
  movel([0.314880, -1.385235, -2.546069, -0.781086, 1.570796, 1.885677],accel_mss,speed_ms,0,blend_radius_m)
  movel([0.314941, -1.384958, -2.546267, -0.781163, 1.570796, 1.885737],accel_mss,speed_ms,0,blend_radius_m)
  movel([0.315016, -1.384678, -2.546469, -0.781242, 1.570796, 1.885812],accel_mss,speed_ms,0,blend_radius_m)
  movel([0.315112, -1.384396, -2.546671, -0.781322, 1.570796, 1.885909],accel_mss,speed_ms,0,blend_radius_m)
  movel([0.315224, -1.384115, -2.546873, -0.781401, 1.570796, 1.886021],accel_mss,speed_ms,0,blend_radius_m)
  movel([0.315355, -1.383832, -2.547076, -0.781481, 1.570796, 1.886151],accel_mss,speed_ms,0,blend_radius_m)
  movel([0.315501, -1.383550, -2.547278, -0.781561, 1.570796, 1.886297],accel_mss,speed_ms,0,blend_radius_m)
  movel([0.315663, -1.383268, -2.547480, -0.781641, 1.570796, 1.886459],accel_mss,speed_ms,0,blend_radius_m)
  movel([0.315841, -1.382992, -2.547678, -0.781719, 1.570796, 1.886637],accel_mss,speed_ms,0,blend_radius_m)
  movel([0.316035, -1.382716, -2.547875, -0.781798, 1.570796, 1.886831],accel_mss,speed_ms,0,blend_radius_m)
  movel([0.316242, -1.382447, -2.548067, -0.781874, 1.570796, 1.887039],accel_mss,speed_ms,0,blend_radius_m)
  movel([0.316464, -1.382184, -2.548255, -0.781949, 1.570796, 1.887260],accel_mss,speed_ms,0,blend_radius_m)
  movel([0.316699, -1.381927, -2.548440, -0.782023, 1.570796, 1.887496],accel_mss,speed_ms,0,blend_radius_m)
  movel([0.316945, -1.381679, -2.548617, -0.782094, 1.570796, 1.887742],accel_mss,speed_ms,0,blend_radius_m)
  movel([0.317202, -1.381438, -2.548788, -0.782162, 1.570796, 1.887999],accel_mss,speed_ms,0,blend_radius_m)
  movel([0.317470, -1.381206, -2.548954, -0.782229, 1.570796, 1.888267],accel_mss,speed_ms,0,blend_radius_m)
  movel([0.317748, -1.380985, -2.549111, -0.782292, 1.570796, 1.888544],accel_mss,speed_ms,0,blend_radius_m)
  movel([0.318653, -1.380294, -2.549604, -0.782491, 1.570796, 1.889449],accel_mss,speed_ms,0,blend_radius_m)
  movel([0.318586, -1.379967, -2.549837, -0.782585, 1.570796, 1.889382],accel_mss,speed_ms,0,blend_radius_m)
  movel([0.318515, -1.379567, -2.550122, -0.782701, 1.570796, 1.889311],accel_mss,speed_ms,0,blend_radius_m)
  movel([0.318460, -1.379160, -2.550410, -0.782818, 1.570796, 1.889256],accel_mss,speed_ms,0,blend_radius_m)
  movel([0.318426, -1.378743, -2.550707, -0.782939, 1.570796, 1.889222],accel_mss,speed_ms,0,blend_radius_m)
  movel([0.318372, -1.377731, -2.551425, -0.783234, 1.570796, 1.889168],accel_mss,speed_ms,0,blend_radius_m)
  movel([0.318336, -1.376711, -2.552146, -0.783532, 1.570796, 1.889132],accel_mss,speed_ms,0,blend_radius_m)
  movel([0.318320, -1.375928, -2.552699, -0.783762, 1.570796, 1.889117],accel_mss,speed_ms,0,blend_radius_m)
  movel([0.318313, -1.375140, -2.553255, -0.783994, 1.570796, 1.889109],accel_mss,speed_ms,0,blend_radius_m)
  movel([0.318313, -1.374350, -2.553811, -0.784228, 1.570796, 1.889109],accel_mss,speed_ms,0,blend_radius_m)
  movel([0.318324, -1.373554, -2.554371, -0.784464, 1.570796, 1.889120],accel_mss,speed_ms,0,blend_radius_m)
  movel([0.318345, -1.372754, -2.554933, -0.784702, 1.570796, 1.889141],accel_mss,speed_ms,0,blend_radius_m)
  movel([0.318374, -1.371950, -2.555496, -0.784943, 1.570796, 1.889170],accel_mss,speed_ms,0,blend_radius_m)
  movel([0.318407, -1.370741, -2.556342, -0.785306, 1.570796, 1.889203],accel_mss,speed_ms,0,blend_radius_m)
  movel([0.318408, -1.369541, -2.557179, -0.785669, 1.570796, 1.889205],accel_mss,speed_ms,0,blend_radius_m)
  movel([0.318376, -1.368351, -2.558008, -0.786030, 1.570796, 1.889172],accel_mss,speed_ms,0,blend_radius_m)
  movel([0.318345, -1.367819, -2.558377, -0.786193, 1.570796, 1.889141],accel_mss,speed_ms,0,blend_radius_m)
  movel([0.318291, -1.367298, -2.558739, -0.786352, 1.570796, 1.889087],accel_mss,speed_ms,0,blend_radius_m)
  movel([0.318219, -1.366783, -2.559096, -0.786510, 1.570796, 1.889016],accel_mss,speed_ms,0,blend_radius_m)
  movel([0.318124, -1.366280, -2.559445, -0.786664, 1.570796, 1.888921],accel_mss,speed_ms,0,blend_radius_m)
  movel([0.318008, -1.365786, -2.559787, -0.786817, 1.570796, 1.888805],accel_mss,speed_ms,0,blend_radius_m)
  movel([0.317894, -1.365379, -2.560068, -0.786942, 1.570796, 1.888690],accel_mss,speed_ms,0,blend_radius_m)
  movel([0.317756, -1.364986, -2.560339, -0.787063, 1.570796, 1.888553],accel_mss,speed_ms,0,blend_radius_m)
  movel([0.317597, -1.364608, -2.560600, -0.787180, 1.570796, 1.888394],accel_mss,speed_ms,0,blend_radius_m)
  movel([0.317419, -1.364241, -2.560854, -0.787294, 1.570796, 1.888215],accel_mss,speed_ms,0,blend_radius_m)
  movel([0.317218, -1.363888, -2.561097, -0.787404, 1.570796, 1.888014],accel_mss,speed_ms,0,blend_radius_m)
  movel([0.316998, -1.363553, -2.561328, -0.787508, 1.570796, 1.887794],accel_mss,speed_ms,0,blend_radius_m)
  movel([0.316760, -1.363235, -2.561546, -0.787607, 1.570796, 1.887556],accel_mss,speed_ms,0,blend_radius_m)
  movel([0.316499, -1.362935, -2.561753, -0.787701, 1.570796, 1.887296],accel_mss,speed_ms,0,blend_radius_m)
  movel([0.316220, -1.362650, -2.561949, -0.787790, 1.570796, 1.887016],accel_mss,speed_ms,0,blend_radius_m)
  movel([0.315920, -1.362382, -2.562133, -0.787874, 1.570796, 1.886716],accel_mss,speed_ms,0,blend_radius_m)
  movel([0.315593, -1.362128, -2.562308, -0.787953, 1.570796, 1.886389],accel_mss,speed_ms,0,blend_radius_m)
  movel([0.315243, -1.361896, -2.562467, -0.788026, 1.570796, 1.886040],accel_mss,speed_ms,0,blend_radius_m)
  movel([0.314859, -1.361672, -2.562621, -0.788096, 1.570796, 1.885655],accel_mss,speed_ms,0,blend_radius_m)
  movel([0.314455, -1.361470, -2.562759, -0.788160, 1.570796, 1.885251],accel_mss,speed_ms,0,blend_radius_m)
  movel([0.314040, -1.361293, -2.562880, -0.788215, 1.570796, 1.884837],accel_mss,speed_ms,0,blend_radius_m)
  movel([0.313611, -1.361138, -2.562987, -0.788264, 1.570796, 1.884407],accel_mss,speed_ms,0,blend_radius_m)
  movel([0.313202, -1.361020, -2.563068, -0.788301, 1.570796, 1.883998],accel_mss,speed_ms,0,blend_radius_m)
  movel([0.312777, -1.360925, -2.563133, -0.788331, 1.570796, 1.883574],accel_mss,speed_ms,0,blend_radius_m)
  movel([0.311989, -1.360781, -2.563231, -0.788377, 1.570796, 1.882786],accel_mss,speed_ms,0,blend_radius_m)
  movel([0.311807, -1.361152, -2.562977, -0.788260, 1.570796, 1.882603],accel_mss,speed_ms,0,blend_radius_m)
  movel([0.311579, -1.361646, -2.562638, -0.788104, 1.570796, 1.882375],accel_mss,speed_ms,0,blend_radius_m)
  movel([0.310419, -1.364402, -2.560742, -0.787244, 1.570796, 1.881216],accel_mss,speed_ms,0,blend_radius_m)
  movel([0.310397, -1.364455, -2.560706, -0.787228, 1.570796, 1.881193],accel_mss,speed_ms,0,blend_radius_m)
  movel([0.310359, -1.364508, -2.560670, -0.787212, 1.570796, 1.881155],accel_mss,speed_ms,0,blend_radius_m)
  movel([0.310331, -1.364535, -2.560651, -0.787203, 1.570796, 1.881127],accel_mss,speed_ms,0,blend_radius_m)
  movel([0.310301, -1.364555, -2.560637, -0.787197, 1.570796, 1.881097],accel_mss,speed_ms,0,blend_radius_m)
  movel([0.310269, -1.364570, -2.560627, -0.787192, 1.570796, 1.881065],accel_mss,speed_ms,0,blend_radius_m)
  movel([0.310191, -1.364588, -2.560614, -0.787187, 1.570796, 1.880987],accel_mss,speed_ms,0,blend_radius_m)
  movel([0.310114, -1.364596, -2.560609, -0.787184, 1.570796, 1.880911],accel_mss,speed_ms,0,blend_radius_m)
  movel([0.309806, -1.364599, -2.560606, -0.787183, 1.570796, 1.880603],accel_mss,speed_ms,0,blend_radius_m)
  movel([0.308187, -1.364604, -2.560603, -0.787182, 1.570796, 1.878983],accel_mss,speed_ms,0,blend_radius_m)
  movel([0.307980, -1.364655, -2.560568, -0.787166, 1.570796, 1.878777],accel_mss,speed_ms,0,blend_radius_m)
  movel([0.307917, -1.364699, -2.560537, -0.787152, 1.570796, 1.878713],accel_mss,speed_ms,0,blend_radius_m)
  movel([0.307876, -1.364761, -2.560495, -0.787133, 1.570796, 1.878672],accel_mss,speed_ms,0,blend_radius_m)
  movel([0.307833, -1.364876, -2.560416, -0.787098, 1.570796, 1.878630],accel_mss,speed_ms,0,blend_radius_m)
  movel([0.307776, -1.364992, -2.560336, -0.787062, 1.570796, 1.878572],accel_mss,speed_ms,0,blend_radius_m)
  movel([0.307708, -1.365107, -2.560256, -0.787026, 1.570796, 1.878504],accel_mss,speed_ms,0,blend_radius_m)
  movel([0.307355, -1.365641, -2.559887, -0.786861, 1.570796, 1.878152],accel_mss,speed_ms,0,blend_radius_m)
  movel([0.307002, -1.366173, -2.559519, -0.786697, 1.570796, 1.877798],accel_mss,speed_ms,0,blend_radius_m)
  movel([0.306610, -1.366749, -2.559119, -0.786520, 1.570796, 1.877406],accel_mss,speed_ms,0,blend_radius_m)
  movel([0.306213, -1.367322, -2.558722, -0.786345, 1.570796, 1.877010],accel_mss,speed_ms,0,blend_radius_m)
  movel([0.305840, -1.367846, -2.558359, -0.786184, 1.570796, 1.876636],accel_mss,speed_ms,0,blend_radius_m)
  movel([0.305459, -1.368365, -2.557998, -0.786026, 1.570796, 1.876255],accel_mss,speed_ms,0,blend_radius_m)
  movel([0.305006, -1.368964, -2.557581, -0.785844, 1.570796, 1.875803],accel_mss,speed_ms,0,blend_radius_m)
  movel([0.304543, -1.369555, -2.557170, -0.785665, 1.570796, 1.875339],accel_mss,speed_ms,0,blend_radius_m)
  movel([0.304065, -1.370142, -2.556760, -0.785487, 1.570796, 1.874861],accel_mss,speed_ms,0,blend_radius_m)
  movel([0.303576, -1.370722, -2.556355, -0.785312, 1.570796, 1.874372],accel_mss,speed_ms,0,blend_radius_m)
  movel([0.303074, -1.371293, -2.555956, -0.785140, 1.570796, 1.873871],accel_mss,speed_ms,0,blend_radius_m)
  movel([0.302561, -1.371859, -2.555560, -0.784970, 1.570796, 1.873357],accel_mss,speed_ms,0,blend_radius_m)
  movel([0.302037, -1.372416, -2.555169, -0.784803, 1.570796, 1.872833],accel_mss,speed_ms,0,blend_radius_m)
  movel([0.301499, -1.372969, -2.554782, -0.784638, 1.570796, 1.872296],accel_mss,speed_ms,0,blend_radius_m)
  movel([0.300953, -1.373513, -2.554400, -0.784476, 1.570796, 1.871750],accel_mss,speed_ms,0,blend_radius_m)
  movel([0.300394, -1.374049, -2.554023, -0.784317, 1.570796, 1.871190],accel_mss,speed_ms,0,blend_radius_m)
  movel([0.299830, -1.374574, -2.553653, -0.784161, 1.570796, 1.870626],accel_mss,speed_ms,0,blend_radius_m)
  movel([0.299252, -1.375093, -2.553288, -0.784008, 1.570796, 1.870049],accel_mss,speed_ms,0,blend_radius_m)
  movel([0.298667, -1.375600, -2.552930, -0.783858, 1.570796, 1.869464],accel_mss,speed_ms,0,blend_radius_m)
  movel([0.298075, -1.376098, -2.552579, -0.783712, 1.570796, 1.868871],accel_mss,speed_ms,0,blend_radius_m)
  movel([0.297481, -1.376580, -2.552239, -0.783570, 1.570796, 1.868277],accel_mss,speed_ms,0,blend_radius_m)
  movel([0.296879, -1.377052, -2.551905, -0.783432, 1.570796, 1.867675],accel_mss,speed_ms,0,blend_radius_m)
  movel([0.296270, -1.377512, -2.551579, -0.783298, 1.570796, 1.867066],accel_mss,speed_ms,0,blend_radius_m)
  movel([0.295655, -1.377964, -2.551259, -0.783166, 1.570796, 1.866452],accel_mss,speed_ms,0,blend_radius_m)
  movel([0.295032, -1.378401, -2.550949, -0.783039, 1.570796, 1.865828],accel_mss,speed_ms,0,blend_radius_m)
  movel([0.294405, -1.378828, -2.550647, -0.782915, 1.570796, 1.865202],accel_mss,speed_ms,0,blend_radius_m)
  movel([0.293771, -1.379244, -2.550351, -0.782794, 1.570796, 1.864568],accel_mss,speed_ms,0,blend_radius_m)
  movel([0.293150, -1.379636, -2.550072, -0.782681, 1.570796, 1.863946],accel_mss,speed_ms,0,blend_radius_m)
  movel([0.292523, -1.380013, -2.549804, -0.782572, 1.570796, 1.863319],accel_mss,speed_ms,0,blend_radius_m)
  movel([0.291892, -1.380380, -2.549543, -0.782466, 1.570796, 1.862688],accel_mss,speed_ms,0,blend_radius_m)
  movel([0.291258, -1.380730, -2.549293, -0.782366, 1.570796, 1.862054],accel_mss,speed_ms,0,blend_radius_m)
  movel([0.290619, -1.381068, -2.549052, -0.782269, 1.570796, 1.861415],accel_mss,speed_ms,0,blend_radius_m)
  movel([0.289977, -1.381393, -2.548820, -0.782175, 1.570796, 1.860774],accel_mss,speed_ms,0,blend_radius_m)
  movel([0.289332, -1.381702, -2.548600, -0.782087, 1.570796, 1.860129],accel_mss,speed_ms,0,blend_radius_m)
  movel([0.288727, -1.381980, -2.548401, -0.782007, 1.570796, 1.859523],accel_mss,speed_ms,0,blend_radius_m)
  movel([0.288119, -1.382244, -2.548213, -0.781932, 1.570796, 1.858916],accel_mss,speed_ms,0,blend_radius_m)
  movel([0.287511, -1.382498, -2.548031, -0.781860, 1.570796, 1.858307],accel_mss,speed_ms,0,blend_radius_m)
  movel([0.286902, -1.382737, -2.547861, -0.781792, 1.570796, 1.857699],accel_mss,speed_ms,0,blend_radius_m)
  movel([0.286307, -1.382957, -2.547703, -0.781729, 1.570796, 1.857103],accel_mss,speed_ms,0,blend_radius_m)
  movel([0.285711, -1.383164, -2.547554, -0.781670, 1.570796, 1.856507],accel_mss,speed_ms,0,blend_radius_m)
  movel([0.285117, -1.383359, -2.547415, -0.781615, 1.570796, 1.855913],accel_mss,speed_ms,0,blend_radius_m)
  movel([0.284524, -1.383537, -2.547287, -0.781565, 1.570796, 1.855320],accel_mss,speed_ms,0,blend_radius_m)
  movel([0.283920, -1.383708, -2.547165, -0.781516, 1.570796, 1.854716],accel_mss,speed_ms,0,blend_radius_m)
  movel([0.283316, -1.383862, -2.547055, -0.781473, 1.570796, 1.854113],accel_mss,speed_ms,0,blend_radius_m)
  movel([0.282717, -1.384002, -2.546954, -0.781433, 1.570796, 1.853514],accel_mss,speed_ms,0,blend_radius_m)
  movel([0.282120, -1.384130, -2.546862, -0.781397, 1.570796, 1.852916],accel_mss,speed_ms,0,blend_radius_m)
  movel([0.281491, -1.384250, -2.546776, -0.781363, 1.570796, 1.852288],accel_mss,speed_ms,0,blend_radius_m)
  movel([0.280864, -1.384358, -2.546698, -0.781332, 1.570796, 1.851660],accel_mss,speed_ms,0,blend_radius_m)
  movel([0.280241, -1.384451, -2.546631, -0.781306, 1.570796, 1.851037],accel_mss,speed_ms,0,blend_radius_m)
  movel([0.279621, -1.384534, -2.546572, -0.781283, 1.570796, 1.850418],accel_mss,speed_ms,0,blend_radius_m)
  movel([0.277452, -1.384799, -2.546382, -0.781208, 1.570796, 1.848248],accel_mss,speed_ms,0,blend_radius_m)
  movel([0.277251, -1.385117, -2.546153, -0.781119, 1.570796, 1.848048],accel_mss,speed_ms,0,blend_radius_m)
  movel([0.277203, -1.385187, -2.546103, -0.781099, 1.570796, 1.847999],accel_mss,speed_ms,0,blend_radius_m)
  movel([0.277149, -1.385253, -2.546056, -0.781080, 1.570796, 1.847945],accel_mss,speed_ms,0,blend_radius_m)
  movel([0.277086, -1.385318, -2.546009, -0.781062, 1.570796, 1.847883],accel_mss,speed_ms,0,blend_radius_m)
  movel([0.277022, -1.385374, -2.545968, -0.781046, 1.570796, 1.847818],accel_mss,speed_ms,0,blend_radius_m)
  movel([0.276953, -1.385427, -2.545930, -0.781031, 1.570796, 1.847750],accel_mss,speed_ms,0,blend_radius_m)
  movel([0.276881, -1.385472, -2.545898, -0.781019, 1.570796, 1.847677],accel_mss,speed_ms,0,blend_radius_m)
  movel([0.276811, -1.385508, -2.545872, -0.781009, 1.570796, 1.847608],accel_mss,speed_ms,0,blend_radius_m)
  movel([0.276739, -1.385536, -2.545852, -0.781001, 1.570796, 1.847536],accel_mss,speed_ms,0,blend_radius_m)
  movel([0.276615, -1.385572, -2.545826, -0.780991, 1.570796, 1.847411],accel_mss,speed_ms,0,blend_radius_m)
  movel([0.276493, -1.385595, -2.545810, -0.780984, 1.570796, 1.847289],accel_mss,speed_ms,0,blend_radius_m)
  movel([0.276373, -1.385607, -2.545801, -0.780981, 1.570796, 1.847170],accel_mss,speed_ms,0,blend_radius_m)
  movel([0.273566, -1.385725, -2.545716, -0.780948, 1.570796, 1.844362],accel_mss,speed_ms,0,blend_radius_m)
  movel([0.272276, -1.385778, -2.545678, -0.780933, 1.570796, 1.843072],accel_mss,speed_ms,0,blend_radius_m)
  movel([0.270990, -1.385826, -2.545643, -0.780920, 1.570796, 1.841786],accel_mss,speed_ms,0,blend_radius_m)
  movel([0.270544, -1.385839, -2.545634, -0.780916, 1.570796, 1.841340],accel_mss,speed_ms,0,blend_radius_m)
  movel([0.270100, -1.385843, -2.545631, -0.780915, 1.570796, 1.840897],accel_mss,speed_ms,0,blend_radius_m)
  movel([0.269661, -1.385840, -2.545633, -0.780916, 1.570796, 1.840458],accel_mss,speed_ms,0,blend_radius_m)
  movel([0.269552, -1.385833, -2.545638, -0.780918, 1.570796, 1.840349],accel_mss,speed_ms,0,blend_radius_m)
  movel([0.269447, -1.385814, -2.545652, -0.780923, 1.570796, 1.840243],accel_mss,speed_ms,0,blend_radius_m)
  movel([0.269351, -1.385786, -2.545672, -0.780931, 1.570796, 1.840147],accel_mss,speed_ms,0,blend_radius_m)
  movel([0.269260, -1.385748, -2.545699, -0.780941, 1.570796, 1.840056],accel_mss,speed_ms,0,blend_radius_m)
  movel([0.269200, -1.385705, -2.545731, -0.780954, 1.570796, 1.839996],accel_mss,speed_ms,0,blend_radius_m)
  movel([0.269158, -1.385648, -2.545771, -0.780969, 1.570796, 1.839954],accel_mss,speed_ms,0,blend_radius_m)
  movel([0.269130, -1.385580, -2.545821, -0.780989, 1.570796, 1.839927],accel_mss,speed_ms,0,blend_radius_m)
  movel([0.269124, -1.385500, -2.545878, -0.781011, 1.570796, 1.839921],accel_mss,speed_ms,0,blend_radius_m)
  movel([0.269132, -1.385373, -2.545969, -0.781047, 1.570796, 1.839928],accel_mss,speed_ms,0,blend_radius_m)
  movel([0.269152, -1.385243, -2.546063, -0.781083, 1.570796, 1.839949],accel_mss,speed_ms,0,blend_radius_m)
  movel([0.269185, -1.385110, -2.546159, -0.781121, 1.570796, 1.839981],accel_mss,speed_ms,0,blend_radius_m)
  movel([0.269226, -1.384977, -2.546254, -0.781158, 1.570796, 1.840023],accel_mss,speed_ms,0,blend_radius_m)
  movel([0.269467, -1.384321, -2.546725, -0.781343, 1.570796, 1.840263],accel_mss,speed_ms,0,blend_radius_m)
  movel([0.269717, -1.383666, -2.547195, -0.781528, 1.570796, 1.840513],accel_mss,speed_ms,0,blend_radius_m)
  movel([0.270640, -1.381095, -2.549033, -0.782261, 1.570796, 1.841437],accel_mss,speed_ms,0,blend_radius_m)
  movel([0.269989, -1.381178, -2.548974, -0.782237, 1.570796, 1.840786],accel_mss,speed_ms,0,blend_radius_m)
  movel([0.269338, -1.381260, -2.548915, -0.782213, 1.570796, 1.840134],accel_mss,speed_ms,0,blend_radius_m)
  movel([0.268086, -1.385520, -2.545863, -0.781005, 1.570796, 1.838882],accel_mss,speed_ms,0,blend_radius_m)
  movel([0.267571, -1.387267, -2.544604, -0.780517, 1.570796, 1.838368],accel_mss,speed_ms,0,blend_radius_m)
  movel([0.267049, -1.389011, -2.543343, -0.780035, 1.570796, 1.837846],accel_mss,speed_ms,0,blend_radius_m)
  movel([0.266984, -1.389205, -2.543203, -0.779981, 1.570796, 1.837780],accel_mss,speed_ms,0,blend_radius_m)
  movel([0.266899, -1.389402, -2.543060, -0.779927, 1.570796, 1.837695],accel_mss,speed_ms,0,blend_radius_m)
  movel([0.266802, -1.389596, -2.542920, -0.779874, 1.570796, 1.837598],accel_mss,speed_ms,0,blend_radius_m)
  movel([0.266688, -1.389789, -2.542779, -0.779821, 1.570796, 1.837485],accel_mss,speed_ms,0,blend_radius_m)
  movel([0.266625, -1.389875, -2.542717, -0.779797, 1.570796, 1.837421],accel_mss,speed_ms,0,blend_radius_m)
  movel([0.266549, -1.389957, -2.542658, -0.779775, 1.570796, 1.837345],accel_mss,speed_ms,0,blend_radius_m)
  movel([0.266465, -1.390029, -2.542606, -0.779755, 1.570796, 1.837261],accel_mss,speed_ms,0,blend_radius_m)
  movel([0.266373, -1.390089, -2.542562, -0.779738, 1.570796, 1.837169],accel_mss,speed_ms,0,blend_radius_m)
  movel([0.266275, -1.390139, -2.542525, -0.779725, 1.570796, 1.837071],accel_mss,speed_ms,0,blend_radius_m)
  movel([0.266174, -1.390173, -2.542501, -0.779715, 1.570796, 1.836971],accel_mss,speed_ms,0,blend_radius_m)
  movel([0.265882, -1.390248, -2.542446, -0.779695, 1.570796, 1.836678],accel_mss,speed_ms,0,blend_radius_m)
  movel([0.265592, -1.390312, -2.542400, -0.779677, 1.570796, 1.836388],accel_mss,speed_ms,0,blend_radius_m)
  movel([0.265304, -1.390363, -2.542363, -0.779663, 1.570796, 1.836100],accel_mss,speed_ms,0,blend_radius_m)
  movel([0.265018, -1.390406, -2.542332, -0.779652, 1.570796, 1.835814],accel_mss,speed_ms,0,blend_radius_m)
  movel([0.263787, -1.390563, -2.542218, -0.779609, 1.570796, 1.834583],accel_mss,speed_ms,0,blend_radius_m)
  movel([0.263242, -1.392448, -2.540845, -0.779096, 1.570796, 1.834038],accel_mss,speed_ms,0,blend_radius_m)
  movel([0.262698, -1.394331, -2.539469, -0.778588, 1.570796, 1.833494],accel_mss,speed_ms,0,blend_radius_m)
  movel([0.272703, -1.395923, -2.538303, -0.778164, 1.570796, 1.843499],accel_mss,speed_ms,0,blend_radius_m)
  movel([0.276528, -1.396564, -2.537831, -0.777994, 1.570796, 1.847325],accel_mss,speed_ms,0,blend_radius_m)
  movel([0.282659, -1.397627, -2.537049, -0.777713, 1.570796, 1.853455],accel_mss,speed_ms,0,blend_radius_m)
  movel([0.282853, -1.397644, -2.537037, -0.777708, 1.570796, 1.853649],accel_mss,speed_ms,0,blend_radius_m)
  movel([0.282907, -1.397619, -2.537055, -0.777715, 1.570796, 1.853704],accel_mss,speed_ms,0,blend_radius_m)
  movel([0.283027, -1.397508, -2.537137, -0.777744, 1.570796, 1.853823],accel_mss,speed_ms,0,blend_radius_m)
  movel([0.283179, -1.397290, -2.537297, -0.777802, 1.570796, 1.853976],accel_mss,speed_ms,0,blend_radius_m)
  movel([0.283589, -1.396576, -2.537823, -0.777990, 1.570796, 1.854385],accel_mss,speed_ms,0,blend_radius_m)
  movel([0.283756, -1.396305, -2.538022, -0.778062, 1.570796, 1.854552],accel_mss,speed_ms,0,blend_radius_m)
  movel([0.283903, -1.396083, -2.538185, -0.778121, 1.570796, 1.854699],accel_mss,speed_ms,0,blend_radius_m)
  movel([0.283928, -1.396051, -2.538208, -0.778130, 1.570796, 1.854725],accel_mss,speed_ms,0,blend_radius_m)
  movel([0.283963, -1.396026, -2.538226, -0.778136, 1.570796, 1.854759],accel_mss,speed_ms,0,blend_radius_m)
  movel([0.284043, -1.395984, -2.538257, -0.778147, 1.570796, 1.854840],accel_mss,speed_ms,0,blend_radius_m)
  movel([0.284126, -1.395948, -2.538284, -0.778157, 1.570796, 1.854923],accel_mss,speed_ms,0,blend_radius_m)
  movel([0.284207, -1.395920, -2.538304, -0.778164, 1.570796, 1.855003],accel_mss,speed_ms,0,blend_radius_m)
  movel([0.287616, -1.394952, -2.539014, -0.778422, 1.570796, 1.858413],accel_mss,speed_ms,0,blend_radius_m)
  movel([0.290959, -1.394014, -2.539702, -0.778674, 1.570796, 1.861755],accel_mss,speed_ms,0,blend_radius_m)
  movel([0.291093, -1.393981, -2.539725, -0.778682, 1.570796, 1.861889],accel_mss,speed_ms,0,blend_radius_m)
  movel([0.291227, -1.393955, -2.539745, -0.778689, 1.570796, 1.862023],accel_mss,speed_ms,0,blend_radius_m)
  movel([0.291358, -1.393937, -2.539758, -0.778694, 1.570796, 1.862154],accel_mss,speed_ms,0,blend_radius_m)
  movel([0.291448, -1.393937, -2.539758, -0.778694, 1.570796, 1.862244],accel_mss,speed_ms,0,blend_radius_m)
  movel([0.291528, -1.393954, -2.539745, -0.778690, 1.570796, 1.862324],accel_mss,speed_ms,0,blend_radius_m)
  movel([0.293056, -1.394468, -2.539369, -0.778552, 1.570796, 1.863852],accel_mss,speed_ms,0,blend_radius_m)
  movel([0.293924, -1.394764, -2.539152, -0.778472, 1.570796, 1.864721],accel_mss,speed_ms,0,blend_radius_m)
  movel([0.294788, -1.395066, -2.538931, -0.778392, 1.570796, 1.865584],accel_mss,speed_ms,0,blend_radius_m)
  movel([0.296791, -1.395787, -2.538402, -0.778200, 1.570796, 1.867587],accel_mss,speed_ms,0,blend_radius_m)
  movel([0.301951, -1.397690, -2.537003, -0.777696, 1.570796, 1.872747],accel_mss,speed_ms,0,blend_radius_m)
  movel([0.301718, -1.398099, -2.536701, -0.777589, 1.570796, 1.872514],accel_mss,speed_ms,0,blend_radius_m)
  movel([0.299298, -1.402391, -2.533523, -0.776475, 1.570796, 1.870094],accel_mss,speed_ms,0,blend_radius_m)
  movel([0.298777, -1.403305, -2.532843, -0.776241, 1.570796, 1.869573],accel_mss,speed_ms,0,blend_radius_m)
  movel([0.298313, -1.404115, -2.532240, -0.776035, 1.570796, 1.869110],accel_mss,speed_ms,0,blend_radius_m)
  movel([0.298297, -1.404137, -2.532223, -0.776029, 1.570796, 1.869093],accel_mss,speed_ms,0,blend_radius_m)
  movel([0.298275, -1.404158, -2.532207, -0.776024, 1.570796, 1.869071],accel_mss,speed_ms,0,blend_radius_m)
  movel([0.298254, -1.404168, -2.532200, -0.776021, 1.570796, 1.869050],accel_mss,speed_ms,0,blend_radius_m)
  movel([0.298234, -1.404166, -2.532201, -0.776022, 1.570796, 1.869031],accel_mss,speed_ms,0,blend_radius_m)
  movel([0.297351, -1.403672, -2.532570, -0.776148, 1.570796, 1.868147],accel_mss,speed_ms,0,blend_radius_m)
  movel([0.296363, -1.403113, -2.532986, -0.776290, 1.570796, 1.867159],accel_mss,speed_ms,0,blend_radius_m)
  movel([0.295202, -1.402439, -2.533487, -0.776462, 1.570796, 1.865998],accel_mss,speed_ms,0,blend_radius_m)
  movel([0.293033, -1.401227, -2.534388, -0.776774, 1.570796, 1.863829],accel_mss,speed_ms,0,blend_radius_m)
  movel([0.292106, -1.400758, -2.534736, -0.776895, 1.570796, 1.862902],accel_mss,speed_ms,0,blend_radius_m)
  movel([0.292065, -1.400781, -2.534719, -0.776890, 1.570796, 1.862862],accel_mss,speed_ms,0,blend_radius_m)
  movel([0.291975, -1.400876, -2.534648, -0.776865, 1.570796, 1.862771],accel_mss,speed_ms,0,blend_radius_m)
  movel([0.291907, -1.400979, -2.534572, -0.776838, 1.570796, 1.862703],accel_mss,speed_ms,0,blend_radius_m)
  movel([0.288768, -1.407007, -2.530075, -0.775306, 1.570796, 1.859564],accel_mss,speed_ms,0,blend_radius_m)
  movel([0.288784, -1.407053, -2.530041, -0.775295, 1.570796, 1.859580],accel_mss,speed_ms,0,blend_radius_m)
  movel([0.288827, -1.407064, -2.530033, -0.775292, 1.570796, 1.859623],accel_mss,speed_ms,0,blend_radius_m)
